// TIA Portal project "ปริญญานิพนธ์" (V17)

(* hardware
DEVICE "S7-1500/ET200MP station_1"  S7-1500 station
   slot 0: "Rail_0"  Rack  6ES7 590-1***0-0AA0
   slot 1: "PLC_1"  CPU 1511-1 PN  6ES7 511-1AK02-0AB0  V2.9
      slot 3: "CPU display_1"  6ES7591-1AA00-0AA0
      slot 32768: "PROFINET interface_1"  X1
         slot 32769: "Port_1"  X1 P1
         slot 32770: "Port_2"  X1 P2
      slot 34817: "Virtual CP interface port_1"  Virtual CP interface port  Virtual CP interface port
DEVICE "HMI_1"  TP900 Comfort
   slot 0: "HMI_1"  TP900 Comfort  6AV2 124-0JC01-0AX0  17.0.0.0
   slot 1: "HMI_RT_1"  TP900 Comfort  6AV2 124-0JC01-0AX0  17.0.0.0
   slot 5: "HMI_1.IE_CP_1"  PROFINET Interface  17.0.0.0
      slot 1: "PROFINET Interface_1"  PROFINET Interface
         slot 1: "Port_1"  Port
         slot 2: "Port_2"  Port
   slot 7: "HMI_1.MPI/DP_CP_1"  MPI/DP Interface  17.0.0.0
*)

// ===== PLC "PLC_1"  CPU 1511-1 PN =====

VAR_GLOBAL   // PLC tag table "Default tag table"
   "ยา 1" AT %MW850 : Word;
   "ยา 2" AT %MW852 : Word;
   "ยา 3" AT %MW854 : Word;
   "ยา 4" AT %MW856 : Word;
   "ยา 5" AT %MW858 : Word;
   "ยา 6" AT %MW860 : Word;
   "ยา 7" AT %MW862 : Word;
   "ยา 8" AT %MW864 : Word;
   "ยา 9" AT %MW866 : Word;
   "ยา 10" AT %MW868 : Word;
   "ยา 11" AT %MW870 : Word;
   "ยา 12" AT %MW872 : Word;
   "ยา 13" AT %MW874 : Word;
   "ยา 14" AT %MW876 : Word;
   "ยา 15" AT %MW878 : Word;
   "ยา 16" AT %MW880 : Word;
   "ยา 17" AT %MW882 : Word;
   "ยา 18" AT %MW884 : Word;
   "ยา 19" AT %MW886 : Word;
   "ยา 20" AT %MW888 : Word;
   "ยา 21" AT %MW890 : Word;
   "ยา 22" AT %MW892 : Word;
   "ยา 23" AT %MW894 : Word;
   "ยา 24" AT %MW896 : Word;
   "ยา 25" AT %MW898 : Word;
   "ยา 26" AT %MW900 : Word;
   "ยา 27" AT %MW902 : Word;
   "ยา 28" AT %MW904 : Word;
   "ยา 29" AT %MW906 : Word;
   "ยา 30" AT %MW908 : Word;
   "ยา 31" AT %MW910 : Word;
   "ยา 32" AT %MW912 : Word;
   "ยา 33" AT %MW914 : Word;
   "ยา 34" AT %MW916 : Word;
   "ยา 35" AT %MW918 : Word;
   "ยา 36" AT %MW920 : Word;
   "ยา 37" AT %MW922 : Word;
   "ยา 38" AT %MW924 : Word;
   "ยา 39" AT %MW926 : Word;
   "ยา 40" AT %MW928 : Word;
   "ยา 41" AT %MW930 : Word;
   "ยา 42" AT %MW932 : Word;
   "ยา 43" AT %MW934 : Word;
   "ยา 44" AT %MW936 : Word;
   "ยา 45" AT %MW938 : Word;
   "ยา 46" AT %MW940 : Word;
   "ยา 47" AT %MW942 : Word;
   "ยา 48" AT %MW944 : Word;
   "ยา 49" AT %MW946 : Word;
   "ยา 50" AT %MW948 : Word;
   "ยา 51" AT %MW950 : Word;
   "ยา 52" AT %MW952 : Word;
   "ยา 53" AT %MW954 : Word;
   "ยา 54" AT %MW956 : Word;
   "ยา 55" AT %MW958 : Word;
   "ยา 56" AT %MW960 : Word;
   "ยา 57" AT %MW962 : Word;
   "ยา 58" AT %MW964 : Word;
   "ยา 59" AT %MW966 : Word;
   "ยา 60" AT %MW968 : Word;
   "ยา 61" AT %MW970 : Word;
   "ยา 62" AT %MW972 : Word;
   "ยา 63" AT %MW974 : Word;
   "ยา 64" AT %MW976 : Word;
   "ยา 65" AT %MW978 : Word;
   "ยา 66" AT %MW980 : Word;
   "ยา 67" AT %MW982 : Word;
   "ยา 68" AT %MW984 : Word;
   "ยา 69" AT %MW986 : Word;
   "ยา 70" AT %MW988 : Word;
   "ยา 71" AT %MW990 : Word;
   "ยา 72" AT %MW992 : Word;
   "ยา 73" AT %MW994 : Word;
   "ยา 74" AT %MW996 : Word;
   "ยา 75" AT %MW998 : Word;
   "ยา 76" AT %MW1000 : Word;
   "ยา 77" AT %MW1002 : Word;
   "ยา 78" AT %MW1004 : Word;
   "ยา 79" AT %MW1006 : Word;
   "ยา 80" AT %MW1008 : Word;
   "ยา 81" AT %MW1010 : Word;
   "ยา 82" AT %MW1012 : Word;
   "ยา 83" AT %MW1014 : Word;
   "ยา 84" AT %MW1016 : Word;
   "ยา 85" AT %MW1018 : Word;
   "ยา 86" AT %MW1020 : Word;
   "ยา 87" AT %MW1022 : Word;
   "ยา 88" AT %MW1024 : Word;
   "ยา 89" AT %MW1026 : Word;
   "ยา 90" AT %MW1028 : Word;
   "ยา 91" AT %MW1030 : Word;
   "ยา 92" AT %MW1032 : Word;
   "ยา 93" AT %MW1034 : Word;
   "ยา 94" AT %MW1036 : Word;
   "ยา 95" AT %MW1038 : Word;
   "ยา 96" AT %MW1040 : Word;
   "ยา 97" AT %MW1042 : Word;
   "ยา 98" AT %MW1044 : Word;
   "ยา 99" AT %MW1046 : Word;
   "ยา 100" AT %MW1048 : Word;
   "ยา 101" AT %MW1050 : Word;
   "ยา 102" AT %MW1052 : Word;
   "ยา 103" AT %MW1054 : Word;
   "ยา 104" AT %MW1056 : Word;
   "ยา 105" AT %MW1058 : Word;
   "ยา 106" AT %MW1060 : Word;
   "ยา 107" AT %MW1062 : Word;
   "ยา 108" AT %MW1064 : Word;
   "ยา 109" AT %MW1066 : Word;
   "ยา 110" AT %MW1068 : Word;
   "ยา 111" AT %MW1070 : Word;
   "ยา 112" AT %MW1072 : Word;
   "ยา 113" AT %MW1074 : Word;
   "ยา 114" AT %MW1076 : Word;
   "ยา 115" AT %MW1078 : Word;
   "ยา 116" AT %MW1080 : Word;
   "ยา 117" AT %MW1082 : Word;
   "ยา 118" AT %MW1084 : Word;
   "ยา 119" AT %MW1086 : Word;
   "ยา 120" AT %MW1088 : Word;
   "ยา 121" AT %MW1090 : Word;
   "ยา 122" AT %MW1092 : Word;
   "ยา 123" AT %MW1094 : Word;
   "ยา 124" AT %MW1096 : Word;
   "ยา 125" AT %MW1098 : Word;
   "ยา 126" AT %MW1100 : Word;
   "ยา 127" AT %MW1102 : Word;
   "ยา 128" AT %MW1104 : Word;
   "ยา 129" AT %MW1106 : Word;
   "ยา 130" AT %MW1108 : Word;
   "ยา 131" AT %MW1110 : Word;
   "ยา 132" AT %MW1112 : Word;
   "ยา 133" AT %MW1114 : Word;
   "ยา 134" AT %MW1116 : Word;
   "ยา 135" AT %MW1118 : Word;
   "ยา 136" AT %MW1120 : Word;
   "ยา 137" AT %MW1122 : Word;
   "ยา 138" AT %MW1124 : Word;
   "ยา 139" AT %MW1126 : Word;
   "ยา 140" AT %MW1128 : Word;
   "ยา 141" AT %MW1130 : Word;
   "ยา 142" AT %MW1132 : Word;
   "ยา 143" AT %MW1134 : Word;
   "ยา 144" AT %MW1136 : Word;
   "ยา 145" AT %MW1138 : Word;
   "ยา 146" AT %MW1140 : Word;
   "ยา 147" AT %MW1142 : Word;
   "ยา 148" AT %MW1144 : Word;
   "ยา 149" AT %MW1146 : Word;
   "ยา 150" AT %MW1148 : Word;
   "ยา 151" AT %MW1150 : Word;
   "ยา 152" AT %MW1152 : Word;
   "ยา 153" AT %MW1154 : Word;
   "ยา 154" AT %MW1156 : Word;
   "ยา 155" AT %MW1158 : Word;
   "ยา 156" AT %MW1160 : Word;
   "ยา 157" AT %MW1162 : Word;
   "ยา 158" AT %MW1164 : Word;
   "ยา 159" AT %MW1166 : Word;
   "ยา 160" AT %MW1168 : Word;
   "ยา 161" AT %MW1170 : Word;
   "ยา 162" AT %MW1172 : Word;
   "ยา 163" AT %MW1174 : Word;
   "\ยา 164" AT %MW1176 : Word;
   "ยา 165" AT %MW1178 : Word;
   "ยา 166" AT %MW1180 : Word;
   "ยา 167" AT %MW1182 : Word;
   "ยา 168" AT %MW1184 : Word;
   "ยา 169" AT %MW1186 : Word;
   "ยา 170" AT %MW1188 : Word;
   "ยา 171" AT %MW1190 : Word;
   "ยา 172" AT %MW1192 : Word;
   "ยา 173" AT %MW1194 : Word;
   "ยา 174" AT %MW1196 : Word;
   "ยา 175" AT %MW1198 : Word;
   "ยา 176" AT %MW1200 : Word;
   "ยา 177" AT %MW1202 : Word;
   "ยา 178" AT %MW1204 : Word;
   "ยา 179" AT %MW1206 : Word;
   "ยา 180" AT %MW1208 : Word;
   "ยา 181" AT %MW1210 : Word;
   "ยา 182" AT %MW1212 : Word;
   "ยา 183" AT %MW1214 : Word;
   "ยา 184" AT %MW1216 : Word;
   "ยา 185" AT %MW1218 : Word;
   "ยา 186" AT %MW1220 : Word;
   "ยา 187" AT %MW1222 : Word;
   "ยา 188" AT %MW1224 : Word;
   "ยา 189" AT %MW1226 : Word;
   "ยา 190" AT %MW1228 : Word;
   "ยา 191" AT %MW1230 : Word;
   "ยา 192" AT %MW1232 : Word;
   "ยา 193" AT %MW1234 : Word;
   "ยา 194" AT %MW1236 : Word;
   "ยา 195" AT %MW1238 : Word;
   "ยา 196" AT %MW1240 : Word;
   "ยา 197" AT %MW1242 : Word;
   "ยา 198" AT %MW1244 : Word;
   "ยา 199" AT %MW1246 : Word;
   "ยา 200" AT %MW1248 : Word;
   "ยา 201" AT %MW1250 : Word;
   "ยา 202" AT %MW1252 : Word;
   "ยา 203" AT %MW1254 : Word;
   "ยา 204" AT %MW1256 : Word;
   "ยา 205" AT %MW1258 : Word;
   "ยา 206" AT %MW1260 : Word;
   "ยา 207" AT %MW1262 : Word;
   "ยา 208" AT %MW1264 : Word;
   "ยา 209" AT %MW1266 : Word;
   "ยา 210" AT %MW1268 : Word;
   "ยา 211" AT %MW1270 : Word;
   "ยา 212" AT %MW1272 : Word;
   "ยา 213" AT %MW1274 : Word;
   "ยา 214" AT %MW1276 : Word;
   "ยา 215" AT %MW1278 : Word;
   "ยา 216" AT %MW1280 : Word;
   "ยา 217" AT %MW1282 : Word;
   "ยา 218" AT %MW1284 : Word;
   "ยา 219" AT %MW1286 : Word;
   "ยา 220" AT %MW1288 : Word;
   "ยา 221" AT %MW1290 : Word;
   "ยา 222" AT %MW1292 : Word;
   "ยา 223" AT %MW1294 : Word;
   "ยา 224" AT %MW1296 : Word;
   "ยา 225" AT %MW1298 : Word;
   "ยา 226" AT %MW1300 : Word;
   "ยา 227" AT %MW1302 : Word;
   "ยา 228" AT %MW1304 : Word;
   "ยา 229" AT %MW1306 : Word;
   "ยา 230" AT %MW1308 : Word;
   "ยา 231" AT %MW1310 : Word;
   "ยา 232" AT %MW1312 : Word;
   "ยา 233" AT %MW1314 : Word;
   "ยา 234" AT %MW1316 : Word;
   "ยา 235" AT %MW1318 : Word;
   "ยา 236" AT %MW1320 : Word;
   "ยา 237" AT %MW1322 : Word;
   "ยา 238" AT %MW1324 : Word;
   "ยา 239" AT %MW1326 : Word;
   "ยา 240" AT %MW1328 : Word;
   "ยา 241" AT %MW1330 : Word;
   "ยา 242" AT %MW1332 : Word;
   "ยา 243" AT %MW1334 : Word;
   "ยา 244" AT %MW1336 : Word;
   "ยา 245" AT %MW1338 : Word;
   "ยา 246" AT %MW1340 : Word;
   "ยา 247" AT %MW1342 : Word;
   "ยา 248" AT %MW1344 : Word;
   "ยา 249" AT %MW1346 : Word;
   "ยา 250" AT %MW1348 : Word;
   "ยา 251" AT %MW1350 : Word;
   "ยา 252" AT %MW1352 : Word;
   "ยา 253" AT %MW1354 : Word;
   "ยา 254" AT %MW1356 : Word;
   "ยา 255" AT %MW1358 : Word;
   "ยา 256" AT %MW1360 : Word;
   "ยา 257" AT %MW1362 : Word;
   "ยา 258" AT %MW1364 : Word;
   "ยา 259" AT %MW1366 : Word;
   "ยา 260" AT %MW1368 : Word;
   "ยา 261" AT %MW1370 : Word;
   "ยา 262" AT %MW1372 : Word;
   "ยา 263" AT %MW1374 : Word;
   "ยา 264" AT %MW1376 : Word;
   "ยา 265" AT %MW1378 : Word;
   "ยา 266" AT %MW1380 : Word;
   "ยา 267" AT %MW1382 : Word;
   "ยา 268" AT %MW1384 : Word;
   "ยา 269" AT %MW1386 : Word;
   "ยา 270" AT %MW1388 : Word;
   "ยา 271" AT %MW1390 : Word;
   "ยา 272" AT %MW1392 : Word;
   "ยา 273" AT %MW1394 : Word;
   "ยา 274" AT %MW1396 : Word;
   "ยา 275" AT %MW1398 : Word;
   "ยา 276" AT %MW1400 : Word;
   "ยา 277" AT %MW1402 : Word;
   "ยา 278" AT %MW1404 : Word;
   "ยา 279" AT %MW1406 : Word;
   "ยา 280" AT %MW1408 : Word;
   "ยา 281" AT %MW1410 : Word;
   "ยา 282" AT %MW1412 : Word;
   "ยา 283" AT %MW1414 : Word;
   "ยา 284" AT %MW1416 : Word;
   "ยา 285" AT %MW1418 : Word;
   "ยา 286" AT %MW1420 : Word;
   "ยา 287" AT %MW1422 : Word;
   "ยา 288" AT %MW1424 : Word;
   "ยา 289" AT %MW1426 : Word;
   "ยา 290" AT %MW1428 : Word;
   "ยา 291" AT %MW1430 : Word;
   "ยา 292" AT %MW1432 : Word;
   "ยา 293" AT %MW1434 : Word;
   "ยา 294" AT %MW1436 : Word;
   "ยา 295" AT %MW1438 : Word;
   "ยา 296" AT %MW1440 : Word;
   "ยา 297" AT %MW1442 : Word;
   "ยา 298" AT %MW1444 : Word;
   "ยา 299" AT %MW1446 : Word;
   "ยา 300" AT %MW1448 : Word;
   "ยา 301" AT %MW1450 : Word;
   "ยา 302" AT %MW1452 : Word;
   "ยา 303" AT %MW1454 : Word;
   "ยา 304" AT %MW1456 : Word;
   "ยา 305" AT %MW1458 : Word;
   "ยา 306" AT %MW1460 : Word;
   "ยา 307" AT %MW1462 : Word;
   "ยา 308" AT %MW1464 : Word;
   "ยา 309" AT %MW1466 : Word;
   "ยา 310" AT %MW1468 : Word;
   "ยา 311" AT %MW1470 : Word;
   "ยา 312" AT %MW1472 : Word;
   "ยา 313" AT %MW1474 : Word;
   "ยา 314" AT %MW1476 : Word;
   "ยา 315" AT %MW1478 : Word;
   "ยา 316" AT %MW1480 : Word;
   "ยา 317" AT %MW1482 : Word;
   "ยา 318" AT %MW1484 : Word;
   "ยา 319" AT %MW1486 : Word;
   "ยา 320" AT %MW1488 : Word;
   "ยา 321" AT %MW1490 : Word;
   "ยา 322" AT %MW1492 : Word;
   "ยา 323" AT %MW1494 : Word;
   "ยา 324" AT %MW1496 : Word;
   "ยา 325" AT %MW1498 : Word;
   "ยา 326" AT %MW1500 : Word;
   "ยา 327" AT %MW1502 : Word;
   "ยา 328" AT %MW1504 : Word;
   "ยา 329" AT %MW1506 : Word;
   "ยา 330" AT %MW1508 : Word;
   "ยา 331" AT %MW1510 : Word;
   "ยา 332" AT %MW1512 : Word;
   "ยา 333" AT %MW1514 : Word;
   "ยา 334" AT %MW1516 : Word;
   "ยา 335" AT %MW1518 : Word;
   "ยา 336" AT %MW1520 : Word;
   "ยา 337" AT %MW1522 : Word;
   "ยา 338" AT %MW1524 : Word;
   "ยา 339" AT %MW1526 : Word;
   "ยา 340" AT %MW1528 : Word;
   "ยา 341" AT %MW1530 : Word;
   "ยา 342" AT %MW1532 : Word;
   "ยา 343" AT %MW1534 : Word;
   "ยา 344" AT %MW1536 : Word;
   "ยา 345" AT %MW1538 : Word;
   "ยา 346" AT %MW1540 : Word;
   "ยา 347" AT %MW1542 : Word;
   "ยา 348" AT %MW1544 : Word;
   "ยา 349" AT %MW1546 : Word;
   "ยา 350" AT %MW1548 : Word;
   "ยา 351" AT %MW1550 : Word;
   "ยา 352" AT %MW1552 : Word;
   "ยา 353" AT %MW1554 : Word;
   "ยา 354" AT %MW1556 : Word;
   "ยา 355" AT %MW1558 : Word;
   "ยา 356" AT %MW1560 : Word;
   "ยา 357" AT %MW1562 : Word;
   "ยา 358" AT %MW1564 : Word;
   "ยา 359" AT %MW1566 : Word;
   "ยา 360" AT %MW1568 : Word;
   "ยา 361" AT %MW1570 : Word;
   "ยา 362" AT %MW1572 : Word;
   "ยา 363" AT %MW1574 : Word;
   "ยา 364" AT %MW1576 : Word;
   "ยา 365" AT %MW1578 : Word;
   "ยา 366" AT %MW1580 : Word;
   "ยา 367" AT %MW1582 : Word;
   "ยา 368" AT %MW1584 : Word;
   "ยา 369" AT %MW1586 : Word;
   "ยา 370" AT %MW1588 : Word;
   "ยา 371" AT %MW1590 : Word;
   "ยา 372" AT %MW1592 : Word;
   "ยา 373" AT %MW1594 : Word;
   "ยา 374" AT %MW1596 : Word;
   "ยา 375" AT %MW1598 : Word;
   "ยา 376" AT %MW1600 : Word;
   "ยา 377" AT %MW1602 : Word;
   "ยา 378" AT %MW1604 : Word;
   "ยา 379" AT %MW1606 : Word;
   "ยา 380" AT %MW1608 : Word;
   "ยา 381" AT %MW1610 : Word;
   "ยา 382" AT %MW1612 : Word;
   "ยา 383" AT %MW1614 : Word;
   "ยา 384" AT %MW1616 : Word;
   "ยา 385" AT %MW1618 : Word;
   "ยา 386" AT %MW1620 : Word;
   "ยา 387" AT %MW1622 : Word;
   "ยา 388" AT %MW1624 : Word;
   "ยา 389" AT %MW1626 : Word;
   "ยา 390" AT %MW1628 : Word;
   "ยา 391" AT %MW1630 : Word;
   "ยา 392" AT %MW1632 : Word;
   "ยา 393" AT %MW1634 : Word;
   "ยา 394" AT %MW1636 : Word;
   "ยา 395" AT %MW1638 : Word;
   "ยา 396" AT %MW1640 : Word;
   "ยา 397" AT %MW1642 : Word;
   "ยา 398" AT %MW1644 : Word;
   "ยา 399" AT %MW1646 : Word;
   "ยา 400" AT %MW1648 : Word;
   "ยา 401" AT %MW1650 : Word;
   "ยา 402" AT %MW1652 : Word;
   "ยา 403" AT %MW1654 : Word;
   "ยา 404" AT %MW1656 : Word;
   "ยา 405" AT %MW1658 : Word;
   "ยา 406" AT %MW1660 : Word;
   "ยา 407" AT %MW1662 : Word;
   "ยา 408" AT %MW1664 : Word;
   "ยา 409" AT %MW1666 : Word;
   "ยา 410" AT %MW1668 : Word;
   "ยา 411" AT %MW1670 : Word;
   "ยา 412" AT %MW1672 : Word;
   "ยา 413" AT %MW1674 : Word;
   "ยา 414" AT %MW1676 : Word;
   "ยา 415" AT %MW1678 : Word;
   "ยา 416" AT %MW1680 : Word;
   "ยา 417" AT %MW1682 : Word;
   "ยา 418" AT %MW1684 : Word;
   "ยา 419" AT %MW1686 : Word;
   "ยา 420" AT %MW1688 : Word;
   "ยา 421" AT %MW1690 : Word;
   "ยา 422" AT %MW1692 : Word;
   "ยา 423" AT %MW1694 : Word;
   "ยา 424" AT %MW1696 : Word;
   "ยา 425" AT %MW1698 : Word;
   "ยา 426" AT %MW1700 : Word;
   "ยา 427" AT %MW1702 : Word;
   "ยา 428" AT %MW1704 : Word;
   "ยา 429" AT %MW1706 : Word;
   "ยา 430" AT %MW1708 : Word;
   "ยา 431" AT %MW1710 : Word;
   "ยา 432" AT %MW1712 : Word;
   "ยา 433" AT %MW1714 : Word;
   "ยา 434" AT %MW1716 : Word;
   "ยา 435" AT %MW1718 : Word;
   "ยา 436" AT %MW1720 : Word;
   "ยา 437" AT %MW1722 : Word;
   "ยา 438" AT %MW1724 : Word;
   "ยา 439" AT %MW1726 : Word;
   "ยา 440" AT %MW1728 : Word;
   "ยา 441" AT %MW1730 : Word;
   "ยา 442" AT %MW1732 : Word;
   "ยา 443" AT %MW1734 : Word;
   "ยา 444" AT %MW1736 : Word;
   "ยา 445" AT %MW1738 : Word;
   "ยา 446" AT %MW1740 : Word;
   "ยา 447" AT %MW1742 : Word;
   "ยา 448" AT %MW1744 : Word;
   "ยา 449" AT %MW1746 : Word;
   "ยา 450" AT %MW1748 : Word;
   "ยา 451" AT %MW1750 : Word;
   "ยา 452" AT %MW1752 : Word;
   "ยา 453" AT %MW1754 : Word;
   "ยา 454" AT %MW1756 : Word;
   "ยา 455" AT %MW1758 : Word;
   "ยา 456" AT %MW1760 : Word;
   "ยา 457" AT %MW1762 : Word;
   "ยา 458" AT %MW1764 : Word;
   "ยา 459" AT %MW1766 : Word;
   "ยา 460" AT %MW1768 : Word;
   "ยา 461" AT %MW1770 : Word;
   "ยา 462" AT %MW1772 : Word;
   "ยา 463" AT %MW1774 : Word;
   "ยา 464" AT %MW1776 : Word;
   "ยา 465" AT %MW1778 : Word;
   "ยา 466" AT %MW1780 : Word;
   "ยา 467" AT %MW1782 : Word;
   "ยา 468" AT %MW1784 : Word;
   "ยา 469" AT %MW1786 : Word;
   "ยา 470" AT %MW1788 : Word;
   "ยา 471" AT %MW1790 : Word;
   "ยา 472" AT %MW1792 : Word;
   "ยา 473" AT %MW1794 : Word;
   "ยา 474" AT %MW1796 : Word;
   "ยา 475" AT %MW1798 : Word;
   "ยา 476" AT %MW1800 : Word;
   "ยา 477" AT %MW1802 : Word;
   "ยา 478" AT %MW1804 : Word;
   "ยา 479" AT %MW1806 : Word;
   "ยา 480" AT %MW1808 : Word;
   "ยา 481" AT %MW1810 : Word;
   "ยา 482" AT %MW1812 : Word;
   "ยา 483" AT %MW1814 : Word;
   "ยา 484" AT %MW1816 : Word;
   "ยา 485" AT %MW1818 : Word;
   "ยา 486" AT %MW1820 : Word;
   "ยา 487" AT %MW1822 : Word;
   "ยา 488" AT %MW1824 : Word;
   "ยา 489" AT %MW1826 : Word;
   "ยา 490" AT %MW1828 : Word;
   "ยา 491" AT %MW1830 : Word;
   "ยา 492" AT %MW1832 : Word;
   "ยา 493" AT %MW1834 : Word;
   "ยา 494" AT %MW1836 : Word;
   "ยา 495" AT %MW1838 : Word;
   "ยา 496" AT %MW1840 : Word;
   "ยา 497" AT %MW1842 : Word;
   "ยา 498" AT %MW1844 : Word;
   "ยา 499" AT %MW1846 : Word;
   "ยา 500" AT %MW1848 : Word;
   "ยา 501" AT %MW1850 : Word;
   "ยา 502" AT %MW1852 : Word;
   "ยา 503" AT %MW1854 : Word;
   "ยา 504" AT %MW1856 : Word;
   "ยา 505" AT %MW1858 : Word;
   "ยา 506" AT %MW1860 : Word;
   "ยา 507" AT %MW1862 : Word;
   "ยา 508" AT %MW1864 : Word;
   "ยา 509" AT %MW1866 : Word;
   "ยา 510" AT %MW1868 : Word;
   "ยา 511" AT %MW1870 : Word;
   "ยา 512" AT %MW1872 : Word;
   "ยา 513" AT %MW1874 : Word;
   "ยา 514" AT %MW1876 : Word;
   "ยา 515" AT %MW1878 : Word;
   "ยา 516" AT %MW1880 : Word;
   "ยา 517" AT %MW1882 : Word;
   "ยา 518" AT %MW1884 : Word;
   "ยา 519" AT %MW1886 : Word;
   "ยา 520" AT %MW1888 : Word;
   "ยา 164" AT %MW1890 : Word;
   "แสดงชื่อยา2" AT %MW3044 : Word;
   "จัดเก็บ Servo DATA 1,2" AT %MW3046 : Word;
   "จัดเก็บ Servo DATA 3" AT %MW3048 : Word;
   "เบิกจ่าย Servo DATA 1,2" AT %MW3050 : Word;
   "เบิกจ่าย Servo DATA 3" AT %MW3052 : Word;
   "Output ปุ่มยืนยันหน้า Screen" AT %M1965.1 : Bool;
   "Output Motor 1,2 fower จัดเก็บ 1" AT %M1892.0 : Bool;
   "Output Motor No3 จัดเก็บ 1" AT %M1892.1 : Bool;
   "หยุดโชว์สถานะมารับยาซ้ำ" AT %M1892.2 : Bool;
   "Output Motor No3 จัดเก็บ 2" AT %M1892.3 : Bool;
   "Output Motor No3จัดเก็บ 3" AT %M1892.4 : Bool;
   "Output Motor No3 จัดเก็บ 4" AT %M1892.5 : Bool;
   "Output Motor No3จัดเก็บ 5" AT %M1892.6 : Bool;
   "Output Motor No3 จัดเก็บ 6" AT %M1892.7 : Bool;
   "Output Motor No3 จัดเก็บ 7" AT %M1893.0 : Bool;
   "Output Motor No3 จัดเก็บ 8" AT %M1893.1 : Bool;
   "Output Motor No3 จัดเก็บ 9" AT %M1893.2 : Bool;
   "Output Motor No3 จัดเก็บ10" AT %M1893.3 : Bool;
   "Output Motor No3จัดเก็บ 11" AT %M1893.4 : Bool;
   "Output Motor No3 จัดเก็บ 12" AT %M1893.5 : Bool;
   "Output Motor No3จัดเก็บ 13" AT %M1893.6 : Bool;
   "Output Motor No3 จัดเก็บ 14" AT %M1893.7 : Bool;
   "Output Motor No3 จัดเก็บ 15" AT %M1894.0 : Bool;
   "Output Motor No3 จัดเก็บ 16" AT %M1894.1 : Bool;
   "Output Motor No3 จัดเก็บ 17" AT %M1894.2 : Bool;
   "Output Motor No3 จัดเก็บ 18" AT %M1894.3 : Bool;
   "Output Motor No3จัดเก็บ 19" AT %M1894.4 : Bool;
   "Output Motor No3 จัดเก็บ 20" AT %M1894.5 : Bool;
   "Output Motor No3จัดเก็บ 21" AT %M1894.6 : Bool;
   "Output Motor No3 จัดเก็บ 22" AT %M1894.7 : Bool;
   "Output Motor No3 จัดเก็บ 23" AT %M1895.0 : Bool;
   "Output Motor No3จัดเก็บ 24" AT %M1895.1 : Bool;
   "Output Motor No3 จัดเก็บ 25" AT %M1895.2 : Bool;
   "Output Motor No3จัดเก็บ 26" AT %M1895.3 : Bool;
   "Oupput Motor 3 จัดเก็บ RESET" AT %M1895.4 : Bool;
   "Output Reset พิเศษ จัดเก็บบ" AT %M1895.5 : Bool;
   "Output Motor 1,2 fower จัดเก็บ 2" AT %M1895.6 : Bool;
   "Output Motor 1,2 fower จัดเก็บ 3" AT %M1895.7 : Bool;
   "Output Motor 1,2 fower จัดเก็บ 4" AT %M1896.0 : Bool;
   "Output Motor 1,2 fower จัดเก็บ 5" AT %M1896.1 : Bool;
   "Output Motor 1,2 fower จัดเก็บ 6" AT %M1896.2 : Bool;
   "Output Motor 1,2 fower จัดเก็บ 7" AT %M1896.3 : Bool;
   "Output Motor 1,2 fower จัดเก็บ 8" AT %M1896.4 : Bool;
   "Output Motor 1,2 fower จัดเก็บ 9" AT %M1896.5 : Bool;
   "Output Motor 1,2 fower จัดเก็บ 10" AT %M1896.6 : Bool;
   "Output Motor 1,2 fower จัดเก็บ 11" AT %M1896.7 : Bool;
   "Output Motor 1,2 fower จัดเก็บ 12" AT %M1897.0 : Bool;
   "Output Motor 1,2 fower จัดเก็บ 13" AT %M1897.1 : Bool;
   "Output Motor 1,2 fower จัดเก็บ 14" AT %M1897.2 : Bool;
   "Output Motor 1,2 fower จัดเก็บ 15" AT %M1897.3 : Bool;
   "Output Motor 1,2 fower จัดเก็บ 16" AT %M1897.4 : Bool;
   "Output Motor 1,2 fower จัดเก็บ 17" AT %M1897.5 : Bool;
   "Output Motor 1,2 fower จัดเก็บ 18" AT %M1897.6 : Bool;
   "Output Motor 1,2 fower จัดเก็บ 19" AT %M1897.7 : Bool;
   "Output Motor 1,2 fower จัดเก็บ 20" AT %M1898.0 : Bool;
   "Output test1" AT %M1898.1 : Bool;
   "Outputtest2" AT %M1898.2 : Bool;
   "Step Motor 3 forword_NOซ้าย-ขวา" AT %M1898.3 : Bool;
   "SR Test" AT %M1898.4 : Bool;
   "Emergency stop" AT %M1898.5 : Bool;
   "Reset-All System" AT %M1898.6 : Bool;
END_VAR

VAR_GLOBAL   // PLC tag table "Tag table_1"
   "SR Conveyor1" AT %M100.0 : Bool;
   "SR Conveyor2" AT %M100.1 : Bool;
   "มีการปุ่มกดยืนยัน" AT %M100.2 : Bool;
   "Brushless Motor Conveyor ทำงาน" AT %M100.3 : Bool;
   "Photoelectic sensor 3 ตรวจเจอวัตถุ" AT %M100.4 : Bool;
   "OutputหลังPhotoelectic sensor 3 ตรวจเจอวัตถุ" AT %M100.5 : Bool;
END_VAR

VAR_GLOBAL   // PLC tag table "Tag table_2"
   "SR_System_In Motor No.1" AT %M200.0 : Bool;
   "SR_System_In Motor No.1(1)" AT %M200.1 : Bool;
   "SR_System_In Motor No.1(2)" AT %M200.2 : Bool;
   "SR_System_In Motor No.1(3)" AT %M200.3 : Bool;
   "SR_System_In Motor No.1(4)" AT %M200.4 : Bool;
   "SR_System_In Motor No.1(5)" AT %M200.5 : Bool;
   "SR_System_In Motor No.1(6)" AT %M200.6 : Bool;
   "SR_System_In Motor No.1(7)" AT %M200.7 : Bool;
   "SR_System_In Motor No.1(8)" AT %M201.0 : Bool;
   "SR_System_In Motor No.1(9)" AT %M201.1 : Bool;
   "SR_System_In Motor No.1(10)" AT %M201.2 : Bool;
   "SR_System_In Motor No.1(11)" AT %M201.3 : Bool;
   "SR_System_In Motor No.1(12)" AT %M201.4 : Bool;
   "SR_System_In Motor No.1(13)" AT %M201.5 : Bool;
   "SR_System_In Motor No.1(14)" AT %M201.6 : Bool;
   "SR_System_In Motor No.1(15)" AT %M201.7 : Bool;
   "SR_System_In Motor No.1(16)" AT %M202.0 : Bool;
   "SR_System_In Motor No.1(17)" AT %M202.1 : Bool;
   "SR_System_In Motor No.1(18)" AT %M202.2 : Bool;
   "SR_System_In Motor No.1(19)" AT %M202.3 : Bool;
   "SR_System_In Motor No.1(20)" AT %M202.4 : Bool;
   "SR_System_In Motor No.1(21)" AT %M202.5 : Bool;
   "SR_System_In Motor No.1(22)" AT %M202.6 : Bool;
   "SR_System_In Motor No.1(23)" AT %M202.7 : Bool;
   "SR_System_In Motor No.1(24)" AT %M203.0 : Bool;
   "SR_System_In Motor No.1(25)" AT %M203.1 : Bool;
   "SR_System_In Motor No.1(26)" AT %M203.2 : Bool;
   "SR_System_In Motor No.1(27)" AT %M203.3 : Bool;
   "SR_System_In Motor No.1(28)" AT %M203.4 : Bool;
   "SR_System_In Motor No.1(29)" AT %M203.5 : Bool;
   "SR_System_In Motor No.1(30)" AT %M203.6 : Bool;
   "SR_System_In Motor No.1(31)" AT %M203.7 : Bool;
   "SR_System_In Motor No.1(32)" AT %M204.0 : Bool;
   "SR_System_In Motor No.1(33)" AT %M204.1 : Bool;
   "SR_System_In Motor No.1(34)" AT %M204.2 : Bool;
   "SR_System_In Motor No.1(35)" AT %M204.3 : Bool;
   "SR_System_In Motor No.1(36)" AT %M204.4 : Bool;
   "SR_System_In Motor No.1(37)" AT %M204.5 : Bool;
   "SR_System_In Motor No.1(38)" AT %M204.6 : Bool;
   "SR_System_In Motor No.1(39)" AT %M204.7 : Bool;
   "Output Step Motor No.1" AT %M205.0 : Bool;
   "Output Step Motor No.2" AT %M205.1 : Bool;
   "Output Step Motor No.3" AT %M205.2 : Bool;
   "Output Step Motor No.4" AT %M205.3 : Bool;
   "Output Step Motor No.5" AT %M205.4 : Bool;
   "Output Step Motor No.6" AT %M205.5 : Bool;
   "Output Step Motor No.7" AT %M205.6 : Bool;
   "Output Step Motor No.8" AT %M205.7 : Bool;
   "Output Step Motor No.9" AT %M206.0 : Bool;
   "Output Step Motor No.10" AT %M206.1 : Bool;
   "Output Step Motor No.11" AT %M206.2 : Bool;
   "Output Step Motor No.12" AT %M206.3 : Bool;
   "Output Step Motor No.13" AT %M206.4 : Bool;
   "Output Step Motor No.14" AT %M206.5 : Bool;
   "Output Step Motor No.15" AT %M206.6 : Bool;
   "Output Step Motor No.16" AT %M206.7 : Bool;
   "Output Step Motor No.17" AT %M207.0 : Bool;
   "Output Step Motor No.18" AT %M207.1 : Bool;
   "Output Step Motor No.19" AT %M207.2 : Bool;
   "Output Step Motor No.20" AT %M207.3 : Bool;
   "Stepper Motor  ทำงาน" AT %M207.4 : Bool;
   "Stepper Motor No.1 ทำงาน" AT %M207.5 : Bool;
   "Stepper Motor No.2 ทำงาน" AT %M207.6 : Bool;
END_VAR

VAR_GLOBAL   // PLC tag table "Tag table_3"
   "Output Step Motor No.31" AT %M300.0 : Bool;
   "SR_System_In Motor No.3.1" AT %M300.1 : Bool;
   "Stepper Motor 3 ทำงาน" AT %M300.2 : Bool;
   "Stepper Motor No.3 ทำงาน" AT %M300.3 : Bool;
   "Outputพิเศษ" AT %M300.4 : Bool;
   "SR สำหรับสั่ง Motor 3 ต่อ1(1)" AT %M300.6 : Bool;
   "SR สำหรับสั่ง Motor 3 ต่อ1(2)" AT %M300.7 : Bool;
   "SR สำหรับสั่ง Motor 3 ต่อ1(3)" AT %M301.0 : Bool;
   "SR สำหรับสั่ง Motor 3 ต่อ1(4)" AT %M301.1 : Bool;
   "SR สำหรับสั่ง Motor 3 ต่อ1(5)" AT %M301.2 : Bool;
   "SR สำหรับสั่ง Motor 3 ต่อ1(6)" AT %M301.3 : Bool;
   "SR สำหรับสั่ง Motor 3 ต่อ1(7)" AT %M301.4 : Bool;
   "SR สำหรับสั่ง Motor 3 ต่อ1(8)" AT %M301.5 : Bool;
   "SR สำหรับสั่ง Motor 3 ต่อ1(9)" AT %M301.6 : Bool;
   "SR สำหรับสั่ง Motor 3 ต่อ1(10)" AT %M301.7 : Bool;
   "SR สำหรับสั่ง Motor 3 ต่อ1(11)" AT %M302.0 : Bool;
   "SR สำหรับสั่ง Motor 3 ต่อ1(12)" AT %M302.1 : Bool;
   "SR สำหรับสั่ง Motor 3 ต่อ1(13)" AT %M302.2 : Bool;
   "SR สำหรับสั่ง Motor 3 ต่อ1(14)" AT %M302.3 : Bool;
   "SR สำหรับสั่ง Motor 3 ต่อ1(15)" AT %M302.4 : Bool;
   "SR สำหรับสั่ง Motor 3 ต่อ1(16)" AT %M302.5 : Bool;
   "SR สำหรับสั่ง Motor 3 ต่อ1(17)" AT %M302.6 : Bool;
   "SR สำหรับสั่ง Motor 3 ต่อ1(18)" AT %M302.7 : Bool;
   "SR สำหรับสั่ง Motor 3 ต่อ1(19)" AT %M303.0 : Bool;
   "SR สำหรับสั่ง Motor 3 ต่อ1(20)" AT %M303.1 : Bool;
   "SR_System_In Motor No.3.2" AT %M300.5 : Bool;
   "SR_System_In Motor No.3.3" AT %M303.2 : Bool;
   "SR_System_In Motor No.3.4" AT %M303.3 : Bool;
   "SR_System_In Motor No.3.5" AT %M303.4 : Bool;
   "SR_System_In Motor No.3.6" AT %M303.5 : Bool;
   "SR_System_In Motor No.3.7" AT %M303.6 : Bool;
   "SR_System_In Motor No.3.8" AT %M303.7 : Bool;
   "SR_System_In Motor No.3.9" AT %M304.0 : Bool;
   "SR_System_In Motor No.3.10" AT %M304.1 : Bool;
   "SR_System_In Motor No.3.11" AT %M304.2 : Bool;
   "SR_System_In Motor No.3.12" AT %M304.3 : Bool;
   "SR_System_In Motor No.3.13" AT %M304.4 : Bool;
   "SR_System_In Motor No.3.14" AT %M304.5 : Bool;
   "SR_System_In Motor No.3.15" AT %M304.6 : Bool;
   "SR_System_In Motor No.3.16" AT %M304.7 : Bool;
   "SR_System_In Motor No.3.17" AT %M305.0 : Bool;
   "SR_System_In Motor No.3.18" AT %M305.1 : Bool;
   "SR_System_In Motor No.3.19" AT %M305.2 : Bool;
   "SR_System_In Motor No.3.20" AT %M305.3 : Bool;
   "SR_System_In Motor No.3.21" AT %M305.4 : Bool;
   "SR_System_In Motor No.3.22" AT %M305.5 : Bool;
   "SR_System_In Motor No.3.23" AT %M305.6 : Bool;
   "SR_System_In Motor No.3.24" AT %M305.7 : Bool;
   "SR_System_In Motor No.3.25" AT %M306.0 : Bool;
   "SR_System_In Motor No.3.26" AT %M306.1 : Bool;
   "Output Step Motor No.32" AT %M306.2 : Bool;
   "Output Step Motor No.33" AT %M306.3 : Bool;
   "Output Step Motor No.34" AT %M306.4 : Bool;
   "Output Step Motor No.35" AT %M306.5 : Bool;
   "Output Step Motor No.36" AT %M306.6 : Bool;
   "Output Step Motor No.37" AT %M306.7 : Bool;
   "Output Step Motor No.38" AT %M307.0 : Bool;
   "Output Step Motor No.39" AT %M307.1 : Bool;
   "Output Step Motor No.40" AT %M307.2 : Bool;
   "Output Step Motor No.41" AT %M307.3 : Bool;
   "Output Step Motor No.42" AT %M307.4 : Bool;
   "Output Step Motor No.43" AT %M307.5 : Bool;
   "Output Step Motor No.44" AT %M307.6 : Bool;
   "Output Step Motor No.45" AT %M307.7 : Bool;
   "Output Step Motor No.46" AT %M308.0 : Bool;
   "Output Step Motor No.47" AT %M308.1 : Bool;
   "Output Step Motor No.48" AT %M308.2 : Bool;
   "Output Step Motor No.49" AT %M308.3 : Bool;
   "Output Step Motor No.50" AT %M308.4 : Bool;
   "Output Step Motor No.51" AT %M308.5 : Bool;
   "Output Step Motor No.52" AT %M308.6 : Bool;
   "Output Step Motor No.53" AT %M308.7 : Bool;
   "Output Step Motor No.54" AT %M309.0 : Bool;
   "Output Step Motor No.55" AT %M309.1 : Bool;
   "Output Step Motor No.56" AT %M309.2 : Bool;
END_VAR

VAR_GLOBAL   // PLC tag table "Tag table_4"
   "Stepper Motor + Gearhead ทำงาน หมุนไปตำแหน่งเริ่มต้น" AT %M400.0 : Bool;
   "Stepper Motor + Gearhead หยุดทำงาน หมุนไปตำแหน่งเริ่มต้น" AT %M400.1 : Bool;
   "Stepper Motor ทำงาน สไลด์ออก" AT %M400.2 : Bool;
   "Stepper Motor หยุดทำงาน สไลด์ออก" AT %M400.3 : Bool;
   "Stepper Motor ทำงาน หนีบกล่องยา" AT %M400.4 : Bool;
   "Stepper Motor หยุดทำงาน หยุดหนหนีบกล่องยา" AT %M400.5 : Bool;
   "Stepper Motor ทำงาน สไลด์เข้า" AT %M400.6 : Bool;
   "Stepper Motor หยุด ทำงานหยุด สไลด์เข้า" AT %M400.7 : Bool;
   "Stepper Motor + Gearhead ทำงาน หมุนไปตำแหน่งทำงานปล่อยกล่องยาลงบนชั้นเก็บกล่องยา" AT %M401.0 : Bool;
   "Stepper Motor + Gearhead หยุดทำงาน หยุดหมุนไปตำแหน่งทำงานปล่อยกล่องยาลงบนชั้นเก็บกล่องยา" AT %M401.1 : Bool;
   "mmตัดการทำงานครบ 1 รอบ" AT %M401.2 : Bool;
   "Stepper Motor ทำงาน ปล่อยกล่องยา" AT %M401.3 : Bool;
   "Stepper Motor หยุด ทำงาน ปล่อยกล่องยา" AT %M401.4 : Bool;
   "SR Gripper No.1" AT %M401.5 : Bool;
   "SR Gripper No.2" AT %M401.6 : Bool;
   "SR Gripper No.3" AT %M401.7 : Bool;
   "SR Gripper No.4" AT %M402.0 : Bool;
   "SR Gripper No.5" AT %M402.1 : Bool;
   "SR Gripper No.6" AT %M402.2 : Bool;
   "SR Gripper No.7" AT %M402.3 : Bool;
   "SR Gripper No.8" AT %M402.4 : Bool;
   "SR Gripper No.9" AT %M402.5 : Bool;
   "Output เมื่อ Motor ถึงตำแหน่งเป้าหมาย" AT %M402.6 : Bool;
   "output Barcoded" AT %M402.7 : Bool;
   "SR Gripper No.10" AT %M403.0 : Bool;
   "หมุนไปตำแหต่งปล่อยกล่องยา" AT %M403.1 : Bool;
END_VAR

VAR_GLOBAL   // PLC tag table "Tag table_5"
   "Blackword SR(1)" AT %M450.0 : Bool;
   "Blackword SR(2)" AT %M450.1 : Bool;
   "Blackword SR(3)" AT %M450.2 : Bool;
   "Blackword SR(4)" AT %M450.3 : Bool;
   "Stepper Motor Blackword  ทำงาน" AT %M450.4 : Bool;
   "Stepper Motor Blackword No.1 ทำงาน" AT %M450.5 : Bool;
   "Stepper Motor Blackword No.2 ทำงาน" AT %M450.6 : Bool;
   "Output Step Motor Blackword  No.1" AT %M450.7 : Bool;
   "Output Step motor  Backword ทำงาน1" AT %M451.0 : Bool;
   "Output Step Motor Blackword  No.2" AT %M451.1 : Bool;
   "Output Step Motor Blackword  No.3" AT %M451.2 : Bool;
   "Output Step Motor Blackword  No.4" AT %M451.3 : Bool;
   "Output Step Motor Blackword  No.5" AT %M451.4 : Bool;
   "Output Step Motor Blackword  No.6" AT %M451.5 : Bool;
   "Output Step Motor Blackword  No.7" AT %M451.6 : Bool;
   "Output Step Motor Blackword  No.8" AT %M451.7 : Bool;
   "Output Step Motor Blackword  No.9" AT %M452.0 : Bool;
   "Output Step Motor Blackword  No.10" AT %M452.1 : Bool;
   "Output Step Motor Blackword  No.11" AT %M452.2 : Bool;
   "Output Step Motor Blackword  No.12" AT %M452.3 : Bool;
   "Output Step Motor Blackword  No.13" AT %M452.4 : Bool;
   "Output Step Motor Blackword  No.14" AT %M452.5 : Bool;
   "Output Step Motor Blackword  No.15" AT %M452.6 : Bool;
   "Output Step Motor Blackword  No.16" AT %M452.7 : Bool;
   "Output Step Motor Blackword  No.17" AT %M453.0 : Bool;
   "Output Step Motor Blackword  No.18" AT %M453.1 : Bool;
   "Output Step Motor Blackword  No.19" AT %M453.2 : Bool;
   "Output Step Motor Blackword  No.20" AT %M453.3 : Bool;
   "Blackword SR(5)" AT %M453.4 : Bool;
   "Blackword SR(6)" AT %M453.5 : Bool;
   "Blackword SR(7)" AT %M453.6 : Bool;
   "Blackword SR(8)" AT %M453.7 : Bool;
   "Blackword SR(9)" AT %M454.0 : Bool;
   "Blackword SR(10)" AT %M454.1 : Bool;
   "Blackword SR(11)" AT %M454.2 : Bool;
   "Blackword SR(12)" AT %M454.3 : Bool;
   "Blackword SR(13)" AT %M454.4 : Bool;
   "Blackword SR(14)" AT %M454.5 : Bool;
   "Blackword SR(15)" AT %M454.6 : Bool;
   "Blackword SR(16)" AT %M454.7 : Bool;
   "Blackword SR(17)" AT %M455.0 : Bool;
   "Blackword SR(18)" AT %M455.1 : Bool;
   "Blackword SR(19)" AT %M455.2 : Bool;
   "Blackword SR(20)" AT %M455.3 : Bool;
   "Blackword SR(21)" AT %M455.4 : Bool;
   "Blackword SR(22)" AT %M455.5 : Bool;
   "Blackword SR(23)" AT %M455.6 : Bool;
   "Blackword SR(24)" AT %M455.7 : Bool;
   "Blackword SR(25)" AT %M456.0 : Bool;
   "Blackword SR(26)" AT %M456.1 : Bool;
   "Blackword SR(27)" AT %M456.2 : Bool;
   "Blackword SR(28)" AT %M456.3 : Bool;
   "Blackword SR(29)" AT %M456.4 : Bool;
   "Blackword SR(30)" AT %M456.5 : Bool;
   "Blackword SR(31)" AT %M456.6 : Bool;
   "Blackword SR(32)" AT %M456.7 : Bool;
   "Blackword SR(33)" AT %M457.0 : Bool;
   "Blackword SR(34)" AT %M457.1 : Bool;
   "Blackword SR(35)" AT %M457.2 : Bool;
   "Blackword SR(36)" AT %M457.3 : Bool;
   "Blackword SR(37)" AT %M457.4 : Bool;
   "Blackword SR(38)" AT %M457.5 : Bool;
   "Blackword SR(39)" AT %M457.6 : Bool;
   "Blackword SR(40)" AT %M457.7 : Bool;
   "Output Step motor  Backword ทำงาน2" AT %M458.0 : Bool;
   "Output Step motor  Backword ทำงาน3" AT %M458.1 : Bool;
   "Output Step motor  Backword ทำงาน4" AT %M458.2 : Bool;
   "Output Step motor  Backword ทำงาน5" AT %M458.3 : Bool;
   "Output Step motor  Backword ทำงาน6" AT %M458.4 : Bool;
   "Output Step motor  Backword ทำงาน7" AT %M458.5 : Bool;
   "Output Step motor  Backword ทำงาน8" AT %M458.6 : Bool;
   "Output Step motor  Backword ทำงาน9" AT %M458.7 : Bool;
   "Output Step motor  Backword ทำงาน10" AT %M459.0 : Bool;
   "Output Step motor  Backword ทำงาน11" AT %M459.1 : Bool;
   "Output Step motor  Backword ทำงาน12" AT %M459.2 : Bool;
   "Output Step motor  Backword ทำงาน13" AT %M459.3 : Bool;
   "Output Step motor  Backword ทำงาน14" AT %M459.4 : Bool;
   "Output Step motor  Backword ทำงาน15" AT %M459.5 : Bool;
   "Output Step motor  Backword ทำงาน16" AT %M459.6 : Bool;
   "Output Step motor  Backword ทำงาน17" AT %M459.7 : Bool;
   "Output Step motor  Backword ทำงาน18" AT %M460.0 : Bool;
   "Output Step motor  Backword ทำงาน19" AT %M460.1 : Bool;
   "Output Step motor  Backword ทำงาน20" AT %M460.2 : Bool;
END_VAR

VAR_GLOBAL   // PLC tag table "Tag table_6"
   "Output Step Motor Blackword  No.1(1)" AT %M550.0 : Bool;
   "SR Step Motor Blackword 1" AT %M550.1 : Bool;
   "SR Step Motor Blackword 2" AT %M550.2 : Bool;
   "Output test1 พิเศษ" AT %M550.7 : Bool;
   "Stepper Motor Blackword3  ทำงาน" AT %M551.0 : Bool;
   "Stepper Motor Blackword No.3 ทำงาน" AT %M551.1 : Bool;
   "output Step motor  Backword ทำงาน No.3(1)" AT %M551.2 : Bool;
   "Output Step Motor Blackword  No.1(2)" AT %M550.3 : Bool;
   "Output Step Motor Blackword  No.1(3)" AT %M550.4 : Bool;
   "Output Step Motor Blackword  No.1(4)" AT %M550.5 : Bool;
   "Output Step Motor Blackword  No.1(5)" AT %M550.6 : Bool;
   "Output Step Motor Blackword  No.1(6)" AT %M551.3 : Bool;
   "Output Step Motor Blackword  No.1(7)" AT %M551.4 : Bool;
   "Output Step Motor Blackword  No.1(8)" AT %M551.5 : Bool;
   "Output Step Motor Blackword  No.1(9)" AT %M551.6 : Bool;
   "Output Step Motor Blackword  No.1(10)" AT %M551.7 : Bool;
   "Output Step Motor Blackword  No.1(11)" AT %M552.0 : Bool;
   "Output Step Motor Blackword  No.1(12)" AT %M552.1 : Bool;
   "Output Step Motor Blackword  No.1(13)" AT %M552.2 : Bool;
   "Output Step Motor Blackword  No.1(14)" AT %M552.3 : Bool;
   "Output Step Motor Blackword  No.1(15)" AT %M552.4 : Bool;
   "Output Step Motor Blackword  No.1(16)" AT %M552.5 : Bool;
   "Output Step Motor Blackword  No.1(17)" AT %M552.6 : Bool;
   "Output Step Motor Blackword  No.1(18)" AT %M552.7 : Bool;
   "Output Step Motor Blackword  No.1(19)" AT %M553.0 : Bool;
   "Output Step Motor Blackword  No.1(20)" AT %M553.1 : Bool;
   "Output Step Motor Blackword  No.1(21)" AT %M553.2 : Bool;
   "Output Step Motor Blackword  No.1(22)" AT %M553.3 : Bool;
   "Output Step Motor Blackword  No.1(23)" AT %M553.4 : Bool;
   "Output Step Motor Blackword  No.1(24)" AT %M553.5 : Bool;
   "Output Step Motor Blackword  No.1(25)" AT %M553.6 : Bool;
   "Output Step Motor Blackword  No.1(26)" AT %M553.7 : Bool;
   "SR Step Motor Blackword 3" AT %M554.0 : Bool;
   "SR Step Motor Blackword 4" AT %M554.1 : Bool;
   "SR Step Motor Blackword 5" AT %M554.2 : Bool;
   "SR Step Motor Blackword 6" AT %M554.3 : Bool;
   "SR Step Motor Blackword 7" AT %M554.4 : Bool;
   "SR Step Motor Blackword 8" AT %M554.5 : Bool;
   "SR Step Motor Blackword 9" AT %M554.6 : Bool;
   "SR Step Motor Blackword 10" AT %M554.7 : Bool;
   "SR Step Motor Blackword 11" AT %M555.0 : Bool;
   "SR Step Motor Blackword 12" AT %M555.1 : Bool;
   "SR Step Motor Blackword 13" AT %M555.2 : Bool;
   "SR Step Motor Blackword 14" AT %M555.3 : Bool;
   "SR Step Motor Blackword 15" AT %M555.4 : Bool;
   "SR Step Motor Blackword 16" AT %M555.5 : Bool;
   "SR Step Motor Blackword 17" AT %M555.6 : Bool;
   "SR Step Motor Blackword 18" AT %M555.7 : Bool;
   "SR Step Motor Blackword 19" AT %M556.0 : Bool;
   "SR Step Motor Blackword 20" AT %M556.1 : Bool;
   "SR Step Motor Blackword 21" AT %M556.2 : Bool;
   "SR Step Motor Blackword 22" AT %M556.3 : Bool;
   "SR Step Motor Blackword 23" AT %M556.4 : Bool;
   "SR Step Motor Blackword 24" AT %M556.5 : Bool;
   "SR Step Motor Blackword 25" AT %M556.6 : Bool;
   "SR Step Motor Blackword 26" AT %M556.7 : Bool;
   "output Step motor  Backword ทำงาน No.3(2)" AT %M557.0 : Bool;
   "output Step motor  Backword ทำงาน No.3(3)" AT %M557.1 : Bool;
   "output Step motor  Backword ทำงาน No.3(4)" AT %M557.2 : Bool;
   "output Step motor  Backword ทำงาน No.3(5)" AT %M557.3 : Bool;
   "output Step motor  Backword ทำงาน No.3(6)" AT %M557.4 : Bool;
   "output Step motor  Backword ทำงาน No.3(7)" AT %M557.5 : Bool;
   "output Step motor  Backword ทำงาน No.3(8)" AT %M557.6 : Bool;
   "output Step motor  Backword ทำงาน No.3(9)" AT %M557.7 : Bool;
   "output Step motor  Backword ทำงาน No.3(10)" AT %M558.0 : Bool;
   "output Step motor  Backword ทำงาน No.3(11)" AT %M558.1 : Bool;
   "output Step motor  Backword ทำงาน No.3(12)" AT %M558.2 : Bool;
   "output Step motor  Backword ทำงาน No.3(13)" AT %M558.3 : Bool;
   "output Step motor  Backword ทำงาน No.3(14)" AT %M558.4 : Bool;
   "output Step motor  Backword ทำงาน No.3(15)" AT %M558.5 : Bool;
   "output Step motor  Backword ทำงาน No.3(16)" AT %M558.6 : Bool;
   "output Step motor  Backword ทำงาน No.3(17)" AT %M558.7 : Bool;
   "output Step motor  Backword ทำงาน No.3(18)" AT %M559.0 : Bool;
   "output Step motor  Backword ทำงาน No.3(19)" AT %M559.1 : Bool;
   "output Step motor  Backword ทำงาน No.3(20)" AT %M559.2 : Bool;
   "output Step motor  Backword ทำงาน No.3(21)" AT %M559.3 : Bool;
   "output Step motor  Backword ทำงาน No.3(22)" AT %M559.4 : Bool;
   "output Step motor  Backword ทำงาน No.3(23)" AT %M559.5 : Bool;
   "output Step motor  Backword ทำงาน No.3(24)" AT %M559.6 : Bool;
   "output Step motor  Backword ทำงาน No.3(25)" AT %M559.7 : Bool;
   "output Step motor  Backword ทำงาน No.3(26)" AT %M560.0 : Bool;
   "SR Step Motor Blackword 27" AT %M560.1 : Bool;
   "SR Step Motor Blackword 28" AT %M560.2 : Bool;
END_VAR

VAR_GLOBAL   // PLC tag table " เบิกจ่าย Forword"
   "SR Step Motro 1,2  เบิกจ่าย 1" AT %M600.0 : Bool;
   "SR Step Motro 1,2  เบิกจ่าย 2" AT %M600.1 : Bool;
   "SR Step Motro 1,2  เบิกจ่าย 3" AT %M600.2 : Bool;
   "SR Step Motro 1,2  เบิกจ่าย 4" AT %M600.3 : Bool;
   "SR Step Motro 1,2  เบิกจ่าย 5" AT %M600.4 : Bool;
   "SR Step Motro 1,2  เบิกจ่าย 6" AT %M600.5 : Bool;
   "SR Step Motro 1,2  เบิกจ่าย 7" AT %M600.6 : Bool;
   "SR Step Motro 1,2  เบิกจ่าย 8" AT %M600.7 : Bool;
   "SR Step Motro 1,2  เบิกจ่าย 9" AT %M601.0 : Bool;
   "SR Step Motro 1,2  เบิกจ่าย 10" AT %M601.1 : Bool;
   "SR Step Motro 1,2  เบิกจ่าย 11" AT %M601.2 : Bool;
   "SR Step Motro 1,2  เบิกจ่าย 12" AT %M601.3 : Bool;
   "SR Step Motro 1,2  เบิกจ่าย 13" AT %M601.4 : Bool;
   "SR Step Motro 1,2  เบิกจ่าย 14" AT %M601.5 : Bool;
   "SR Step Motro 1,2  เบิกจ่าย 15" AT %M601.6 : Bool;
   "SR Step Motro 1,2  เบิกจ่าย 16" AT %M601.7 : Bool;
   "SR Step Motro 1,2  เบิกจ่าย 17" AT %M602.0 : Bool;
   "SR Step Motro 1,2  เบิกจ่าย 18" AT %M602.1 : Bool;
   "SR Step Motro 1,2  เบิกจ่าย 19" AT %M602.2 : Bool;
   "SR Step Motro 1,2  เบิกจ่าย 20" AT %M602.3 : Bool;
   "Outputเมื่อมีการกดปุ่ม 1" AT %M602.4 : Bool;
   "Outputเมื่อมีการกดปุ่ม 2" AT %M602.5 : Bool;
   "Outputเมื่อมีการกดปุ่ม 3" AT %M602.6 : Bool;
   "Outputเมื่อมีการกดปุ่ม 4" AT %M602.7 : Bool;
   "Outputเมื่อมีการกดปุ่ม 5" AT %M603.0 : Bool;
   "Outputเมื่อมีการกดปุ่ม 6" AT %M603.1 : Bool;
   "Outputเมื่อมีการกดปุ่ม 7" AT %M603.2 : Bool;
   "Outputเมื่อมีการกดปุ่ม 8" AT %M603.3 : Bool;
   "Outputเมื่อมีการกดปุ่ม 9" AT %M603.4 : Bool;
   "Outputเมื่อมีการกดปุ่ม 10" AT %M603.5 : Bool;
   "Outputเมื่อมีการกดปุ่ม 11" AT %M603.6 : Bool;
   "Outputเมื่อมีการกดปุ่ม 12" AT %M603.7 : Bool;
   "Outputเมื่อมีการกดปุ่ม 13" AT %M604.0 : Bool;
   "Outputเมื่อมีการกดปุ่ม 14" AT %M604.1 : Bool;
   "Outputเมื่อมีการกดปุ่ม 15" AT %M604.2 : Bool;
   "Outputเมื่อมีการกดปุ่ม 16" AT %M604.3 : Bool;
   "Outputเมื่อมีการกดปุ่ม 17" AT %M604.4 : Bool;
   "Outputเมื่อมีการกดปุ่ม 18" AT %M604.5 : Bool;
   "Outputเมื่อมีการกดปุ่ม 19" AT %M604.6 : Bool;
   "Outputเมื่อมีการกดปุ่ม 20" AT %M604.7 : Bool;
   "Step motor 1,2 NO" AT %M605.0 : Bool;
   "Step motor 1 NO" AT %M605.1 : Bool;
   "Step motor 2 NO" AT %M605.2 : Bool;
   "Output ทำงานเสด M1,2 forword No.1" AT %M605.3 : Bool;
   "Output ทำงานเสด M1,2 forword No.2" AT %M605.4 : Bool;
   "Output ทำงานเสด M1,2 forword No.3" AT %M605.5 : Bool;
   "Output ทำงานเสด M1,2 forword No.4" AT %M605.6 : Bool;
   "Output ทำงานเสด M1,2 forword No.5" AT %M605.7 : Bool;
   "Output ทำงานเสด M1,2 forword No.6" AT %M606.0 : Bool;
   "Output ทำงานเสด M1,2 forword No.7" AT %M606.1 : Bool;
   "Output ทำงานเสด M1,2 forword No.8" AT %M606.2 : Bool;
   "Output ทำงานเสด M1,2 forword No.9" AT %M606.3 : Bool;
   "Output ทำงานเสด M1,2 forword No.10" AT %M606.4 : Bool;
   "Output ทำงานเสด M1,2 forword No.11" AT %M606.5 : Bool;
   "Output ทำงานเสด M1,2 forword No.12" AT %M606.6 : Bool;
   "Output ทำงานเสด M1,2 forword No.13" AT %M606.7 : Bool;
   "Output ทำงานเสด M1,2 forword No.14" AT %M607.0 : Bool;
   "Output ทำงานเสด M1,2 forword No.15" AT %M607.1 : Bool;
   "Output ทำงานเสด M1,2 forword No.16" AT %M607.2 : Bool;
   "Output ทำงานเสด M1,2 forword No.17" AT %M607.3 : Bool;
   "Output ทำงานเสด M1,2 forword No.18" AT %M607.4 : Bool;
   "Output ทำงานเสด M1,2 forword No.19" AT %M607.5 : Bool;
   "Output ทำงานเสด M1,2 forword No.20" AT %M607.6 : Bool;
END_VAR

VAR_GLOBAL   // PLC tag table " เบิกจ่าย Blackword"
   "SR Step Motro 3  เบิกจ่าย 1" AT %M650.0 : Bool;
   "SR Step Motro 3  เบิกจ่าย 2" AT %M650.1 : Bool;
   "SR Step Motro 3  เบิกจ่าย 3" AT %M650.2 : Bool;
   "SR Step Motro 3  เบิกจ่าย 4" AT %M650.3 : Bool;
   "SR Step Motro 3  เบิกจ่าย 5" AT %M650.4 : Bool;
   "SR Step Motro 3  เบิกจ่าย 6" AT %M650.5 : Bool;
   "SR Step Motro 3  เบิกจ่าย 7" AT %M650.6 : Bool;
   "SR Step Motro 3  เบิกจ่าย 8" AT %M650.7 : Bool;
   "SR Step Motro 3  เบิกจ่าย 9" AT %M651.0 : Bool;
   "SR Step Motro 3  เบิกจ่าย 10" AT %M651.1 : Bool;
   "SR Step Motro 3  เบิกจ่าย 11" AT %M651.2 : Bool;
   "SR Step Motro 3  เบิกจ่าย 12" AT %M651.3 : Bool;
   "SR Step Motro 3  เบิกจ่าย 13" AT %M651.4 : Bool;
   "SR Step Motro 3  เบิกจ่าย 14" AT %M651.5 : Bool;
   "SR Step Motro 3  เบิกจ่าย 15" AT %M651.6 : Bool;
   "SR Step Motro 3  เบิกจ่าย 16" AT %M651.7 : Bool;
   "SR Step Motro 3  เบิกจ่าย 17" AT %M652.0 : Bool;
   "SR Step Motro 3  เบิกจ่าย 18" AT %M652.1 : Bool;
   "SR Step Motro 3  เบิกจ่าย 19" AT %M652.2 : Bool;
   "SR Step Motro 3  เบิกจ่าย 20" AT %M652.3 : Bool;
   "output Step motor No.3  1" AT %M652.4 : Bool;
   "output Step motor No.3  2" AT %M652.5 : Bool;
   "output Step motor No.3  3" AT %M652.6 : Bool;
   "output Step motor No.3  4" AT %M652.7 : Bool;
   "output Step motor No.3  5" AT %M653.0 : Bool;
   "output Step motor No.3  6" AT %M653.1 : Bool;
   "output Step motor No.3  7" AT %M653.2 : Bool;
   "output Step motor No.3  8" AT %M653.3 : Bool;
   "output Step motor No.3  9" AT %M653.4 : Bool;
   "output Step motor No.3  10" AT %M653.5 : Bool;
   "output Step motor No.3  11" AT %M653.6 : Bool;
   "output Step motor No.3  12" AT %M653.7 : Bool;
   "output Step motor No.3  13" AT %M654.0 : Bool;
   "output Step motor No.3  14" AT %M654.1 : Bool;
   "output Step motor No.3  15" AT %M654.2 : Bool;
   "output Step motor No.3  16" AT %M654.3 : Bool;
   "output Step motor No.3  17" AT %M654.4 : Bool;
   "output Step motor No.3  18" AT %M654.5 : Bool;
   "output Step motor No.3  19" AT %M654.6 : Bool;
   "output Step motor No.3  20" AT %M654.7 : Bool;
   "Stepper Motor  ทำงาน Blackword_ON" AT %M655.0 : Bool;
   "Step motor 1 Blackword_NO" AT %M655.1 : Bool;
   "Step motor 2 Blackword_NO" AT %M655.2 : Bool;
   "Output No1,2 Blackword 1" AT %M655.3 : Bool;
   "Output No1,2 Blackword 2" AT %M655.4 : Bool;
   "Output No1,2 Blackword 3" AT %M655.5 : Bool;
   "Output No1,2 Blackword 4" AT %M655.6 : Bool;
   "Output No1,2 Blackword 5" AT %M655.7 : Bool;
   "Output No1,2 Blackword 6" AT %M656.0 : Bool;
   "Output No1,2 Blackword 7" AT %M656.1 : Bool;
   "Output No1,2 Blackword 8" AT %M656.2 : Bool;
   "Output No1,2 Blackword 9" AT %M656.3 : Bool;
   "Output No1,2 Blackword 10" AT %M656.4 : Bool;
   "Output No1,2 Blackword 11" AT %M656.5 : Bool;
   "Output No1,2 Blackword 12" AT %M656.6 : Bool;
   "Output No1,2 Blackword 13" AT %M656.7 : Bool;
   "Output No1,2 Blackword 14" AT %M657.0 : Bool;
   "Output No1,2 Blackword 15" AT %M657.1 : Bool;
   "Output No1,2 Blackword 16" AT %M657.2 : Bool;
   "Output No1,2 Blackword 17" AT %M657.3 : Bool;
   "Output No1,2 Blackword 18" AT %M657.4 : Bool;
   "Output No1,2 Blackword 19" AT %M657.5 : Bool;
   "Output No1,2 Blackword 20" AT %M657.6 : Bool;
END_VAR

VAR_GLOBAL   // PLC tag table "Tag table_7"
   "SR  Gripper เบิกจ่าย 1" AT %M700.0 : Bool;
   "SR  Gripper เบิกจ่าย 2" AT %M700.1 : Bool;
   "Output เวลาหลังจากเคลื่ออนที่ไปถึงตำแหน่งเป้าหมาย" AT %M700.2 : Bool;
   "Stepper Motor ทำงาน สไลด์ ตัวงัดกล่องยาออก" AT %M700.3 : Bool;
   "Stepper Motor หยุดทำงาน หยุดสไลด์ ตัวงัดกล่องยาออก" AT %M700.4 : Bool;
   "Stepper Motor ทำงาน สไลด์ ตัวงัดกล่องยาเข้า" AT %M700.5 : Bool;
   "Stepper Motor หยุดทำงาน หยุดสไลด์ ตัวงัดกล่องยาเข้า" AT %M700.6 : Bool;
   "Stepper Motor ทำงาน สั่งconveyor เคลื่อที่ไปข้างหน้า" AT %M700.7 : Bool;
   "Photoelectic Sensor No.1 เบิกจ่าย" AT %M3600.0 : Bool;
   "Photoelectic Sensor No.2 เบิกจ่าย" AT %M3600.1 : Bool;
   "Photoelectic Sensor No.3 เบิกจ่าย" AT %M3600.2 : Bool;
END_VAR

VAR_GLOBAL   // PLC tag table " เบิกจ่าย Blackword 1"
   "SR Blackword Step motor No.3 เบิกจ่าย 1" AT %M800.0 : Bool;
   "SR Blackword Step motor No.3 เบิกจ่าย 2" AT %M800.1 : Bool;
   "SR Blackword Step motor No.3 เบิกจ่าย 3" AT %M800.2 : Bool;
   "SR Blackword Step motor No.3 เบิกจ่าย 4" AT %M800.3 : Bool;
   "SR Blackword Step motor No.3 เบิกจ่าย 5" AT %M800.4 : Bool;
   "SR Blackword Step motor No.3 เบิกจ่าย 6" AT %M800.5 : Bool;
   "SR Blackword Step motor No.3 เบิกจ่าย 7" AT %M800.6 : Bool;
   "SR Blackword Step motor No.3 เบิกจ่าย 8" AT %M800.7 : Bool;
   "SR Blackword Step motor No.3 เบิกจ่าย 9" AT %M801.0 : Bool;
   "SR Blackword Step motor No.3 เบิกจ่าย 10" AT %M801.1 : Bool;
   "SR Blackword Step motor No.3 เบิกจ่าย 11" AT %M801.2 : Bool;
   "SR Blackword Step motor No.3 เบิกจ่าย 12" AT %M801.3 : Bool;
   "SR Blackword Step motor No.3 เบิกจ่าย 13" AT %M801.4 : Bool;
   "SR Blackword Step motor No.3 เบิกจ่าย 14" AT %M801.5 : Bool;
   "SR Blackword Step motor No.3 เบิกจ่าย 15" AT %M801.6 : Bool;
   "SR Blackword Step motor No.3 เบิกจ่าย 16" AT %M801.7 : Bool;
   "SR Blackword Step motor No.3 เบิกจ่าย 17" AT %M802.0 : Bool;
   "SR Blackword Step motor No.3 เบิกจ่าย 18" AT %M802.1 : Bool;
   "SR Blackword Step motor No.3 เบิกจ่าย 19" AT %M802.2 : Bool;
   "SR Blackword Step motor No.3 เบิกจ่าย 20" AT %M802.3 : Bool;
   "SR Blackword Step motor No.3 เบิกจ่าย 21" AT %M802.4 : Bool;
   "SR Blackword Step motor No.3 เบิกจ่าย 22" AT %M802.5 : Bool;
   "SR Blackword Step motor No.3 เบิกจ่าย 23" AT %M802.6 : Bool;
   "SR Blackword Step motor No.3 เบิกจ่าย 24" AT %M802.7 : Bool;
   "SR Blackword Step motor No.3 เบิกจ่าย 25" AT %M803.0 : Bool;
   "SR Blackword Step motor No.3 เบิกจ่าย 26" AT %M803.1 : Bool;
   "Output Blackword Step motor No.3 เบิกจ่าย 1" AT %M803.2 : Bool;
   "Output Blackword Step motor No.3 เบิกจ่าย 2" AT %M803.3 : Bool;
   "Output Blackword Step motor No.3 เบิกจ่าย 3" AT %M803.4 : Bool;
   "Output Blackword Step motor No.3 เบิกจ่าย 4" AT %M803.5 : Bool;
   "Output Blackword Step motor No.3 เบิกจ่าย 5" AT %M803.6 : Bool;
   "Output Blackword Step motor No.3 เบิกจ่าย 6" AT %M803.7 : Bool;
   "Output Blackword Step motor No.3 เบิกจ่าย 7" AT %M804.0 : Bool;
   "Output Blackword Step motor No.3 เบิกจ่าย 8" AT %M804.1 : Bool;
   "Output Blackword Step motor No.3 เบิกจ่าย 9" AT %M804.2 : Bool;
   "Output Blackword Step motor No.3 เบิกจ่าย 10" AT %M804.3 : Bool;
   "Output Blackword Step motor No.3 เบิกจ่าย 11" AT %M804.4 : Bool;
   "Output Blackword Step motor No.3 เบิกจ่าย 12" AT %M804.5 : Bool;
   "Output Blackword Step motor No.3 เบิกจ่าย 13" AT %M804.6 : Bool;
   "Output Blackword Step motor No.3 เบิกจ่าย 14" AT %M804.7 : Bool;
   "Output Blackword Step motor No.3 เบิกจ่าย 15" AT %M805.0 : Bool;
   "Output Blackword Step motor No.3 เบิกจ่าย 16" AT %M805.1 : Bool;
   "Output Blackword Step motor No.3 เบิกจ่าย 17" AT %M805.2 : Bool;
   "Output Blackword Step motor No.3 เบิกจ่าย 18" AT %M805.3 : Bool;
   "Output Blackword Step motor No.3 เบิกจ่าย 19" AT %M805.4 : Bool;
   "Output Blackword Step motor No.3 เบิกจ่าย 20" AT %M805.5 : Bool;
   "Output Blackword Step motor No.3 เบิกจ่าย 21" AT %M805.6 : Bool;
   "Output Blackword Step motor No.3 เบิกจ่าย 22" AT %M805.7 : Bool;
   "Output Blackword Step motor No.3 เบิกจ่าย 23" AT %M806.0 : Bool;
   "Output Blackword Step motor No.3 เบิกจ่าย 24" AT %M806.1 : Bool;
   "Output Blackword Step motor No.3 เบิกจ่าย 25" AT %M806.2 : Bool;
   "Output Blackword Step motor No.3 เบิกจ่าย 26" AT %M806.3 : Bool;
   "เวลาหลังจากเคลื่อนที่ถึงตำแหน่งเป้าหมาย (26) Blackword" AT %M806.4 : Bool;
   "Step Motor 3 Blackword_NO" AT %M806.5 : Bool;
   "Step Motor No.3 Blackword_NO" AT %M806.6 : Bool;
   "Output black No3 1" AT %M806.7 : Bool;
   "Output black No3 2" AT %M807.0 : Bool;
   "Output black No3 3" AT %M807.1 : Bool;
   "Output black No3 4" AT %M807.2 : Bool;
   "Output black No3 5" AT %M807.3 : Bool;
   "Output black No3 6" AT %M807.4 : Bool;
   "Output black No3 7" AT %M807.5 : Bool;
   "Output black No3 8" AT %M807.6 : Bool;
   "Output black No3 9" AT %M807.7 : Bool;
   "Output black No3 10" AT %M808.0 : Bool;
   "Output black No3 11" AT %M808.1 : Bool;
   "Output black No3 12" AT %M808.2 : Bool;
   "Output black No3 13" AT %M808.3 : Bool;
   "Output black No3 14" AT %M808.4 : Bool;
   "Output black No3 15" AT %M808.5 : Bool;
   "Output black No3 16" AT %M808.6 : Bool;
   "Output black No3 17" AT %M808.7 : Bool;
   "Output black No3 18" AT %M809.0 : Bool;
   "Output black No3 19" AT %M809.1 : Bool;
   "Output black No3 20" AT %M809.2 : Bool;
   "Output black No3 21" AT %M809.3 : Bool;
   "Output black No3 22" AT %M809.4 : Bool;
   "Output black No3 23" AT %M809.5 : Bool;
   "Output black No3 24" AT %M809.6 : Bool;
   "Output black No3 25" AT %M809.7 : Bool;
   "Output black No3 26" AT %M810.0 : Bool;
END_VAR

VAR_GLOBAL   // PLC tag table " เบิกจ่าย Forword 1"
   "SR forword Step motor No.3 เบิกจ่าย 1" AT %M750.0 : Bool;
   "SR forword Step motor No.3 เบิกจ่าย 2" AT %M750.1 : Bool;
   "SR forword Step motor No.3 เบิกจ่าย 3" AT %M750.2 : Bool;
   "SR forword Step motor No.3 เบิกจ่าย 4" AT %M750.3 : Bool;
   "SR forword Step motor No.3 เบิกจ่าย 5" AT %M750.4 : Bool;
   "SR forword Step motor No.3 เบิกจ่าย 6" AT %M750.5 : Bool;
   "SR forword Step motor No.3 เบิกจ่าย 7" AT %M750.6 : Bool;
   "SR forword Step motor No.3 เบิกจ่าย 8" AT %M750.7 : Bool;
   "SR forword Step motor No.3 เบิกจ่าย 9" AT %M751.0 : Bool;
   "SR forword Step motor No.3 เบิกจ่าย 10" AT %M751.1 : Bool;
   "SR forword Step motor No.3 เบิกจ่าย 11" AT %M751.2 : Bool;
   "SR forword Step motor No.3 เบิกจ่าย 12" AT %M751.3 : Bool;
   "SR forword Step motor No.3 เบิกจ่าย 13" AT %M751.4 : Bool;
   "SR forword Step motor No.3 เบิกจ่าย 14" AT %M751.5 : Bool;
   "SR forword Step motor No.3 เบิกจ่าย 15" AT %M751.6 : Bool;
   "SR forword Step motor No.3 เบิกจ่าย 16" AT %M751.7 : Bool;
   "SR forword Step motor No.3 เบิกจ่าย 17" AT %M752.0 : Bool;
   "SR forword Step motor No.3 เบิกจ่าย 18" AT %M752.1 : Bool;
   "SR forword Step motor No.3 เบิกจ่าย 19" AT %M752.2 : Bool;
   "SR forword Step motor No.3 เบิกจ่าย 20" AT %M752.3 : Bool;
   "SR forword Step motor No.3 เบิกจ่าย 21" AT %M752.4 : Bool;
   "SR forword Step motor No.3 เบิกจ่าย 22" AT %M752.5 : Bool;
   "SR forword Step motor No.3 เบิกจ่าย 23" AT %M752.6 : Bool;
   "SR forword Step motor No.3 เบิกจ่าย 24" AT %M752.7 : Bool;
   "SR forword Step motor No.3 เบิกจ่าย 25" AT %M753.0 : Bool;
   "SR forword Step motor No.3 เบิกจ่าย 26" AT %M753.1 : Bool;
   "Output forword Step motor No.3 เบิกจ่าย 1" AT %M753.2 : Bool;
   "Output forword Step motor No.3 เบิกจ่าย 2" AT %M753.3 : Bool;
   "Output forword Step motor No.3 เบิกจ่าย 3" AT %M753.4 : Bool;
   "Output forword Step motor No.3 เบิกจ่าย 4" AT %M753.5 : Bool;
   "Output forword Step motor No.3 เบิกจ่าย 5" AT %M753.6 : Bool;
   "Output forword Step motor No.3 เบิกจ่าย 6" AT %M753.7 : Bool;
   "Output forword Step motor No.3 เบิกจ่าย 7" AT %M754.0 : Bool;
   "Output forword Step motor No.3 เบิกจ่าย 8" AT %M754.1 : Bool;
   "Output forword Step motor No.3 เบิกจ่าย 9" AT %M754.2 : Bool;
   "Output forword Step motor No.3 เบิกจ่าย 10" AT %M754.3 : Bool;
   "Output forword Step motor No.3 เบิกจ่าย 11" AT %M754.4 : Bool;
   "Output forword Step motor No.3 เบิกจ่าย 12" AT %M754.5 : Bool;
   "Output forword Step motor No.3 เบิกจ่าย 13" AT %M754.6 : Bool;
   "Output forword Step motor No.3 เบิกจ่าย 14" AT %M754.7 : Bool;
   "Output forword Step motor No.3 เบิกจ่าย 15" AT %M755.0 : Bool;
   "Output forword Step motor No.3 เบิกจ่าย 16" AT %M755.1 : Bool;
   "Output forword Step motor No.3 เบิกจ่าย 17" AT %M755.2 : Bool;
   "Output forword Step motor No.3 เบิกจ่าย 18" AT %M755.3 : Bool;
   "Output forword Step motor No.3 เบิกจ่าย 19" AT %M755.4 : Bool;
   "Output forword Step motor No.3 เบิกจ่าย 20" AT %M755.5 : Bool;
   "Output forword Step motor No.3 เบิกจ่าย 23" AT %M755.6 : Bool;
   "Output forword Step motor No.3 เบิกจ่าย 24" AT %M755.7 : Bool;
   "Output forword Step motor No.3 เบิกจ่าย 25" AT %M756.0 : Bool;
   "Output forword Step motor No.3 เบิกจ่าย 26" AT %M756.1 : Bool;
   "Output forword Step motor No.3 เบิกจ่าย 21" AT %M756.2 : Bool;
   "Output forword Step motor No.3 เบิกจ่าย 22" AT %M756.3 : Bool;
   "เวลาหลังจากเคลื่อนที่ถึงตำแหน่งเป้าหมาย เบิกจ่าย" AT %M756.4 : Bool;
   "Step Motor 3 forword_NO" AT %M756.5 : Bool;
   "Step Motor No.3 forword_NO" AT %M756.6 : Bool;
   "SR หลังจาก Motor 1,2 ทำงานเสด" AT %M756.7 : Bool;
   "Output ทำงานเสด M 3 forword No.1" AT %M757.0 : Bool;
   "Output ทำงานเสด M 3 forword No.2" AT %M757.1 : Bool;
   "Output ทำงานเสด M 3 forword No.3" AT %M757.2 : Bool;
   "Output ทำงานเสด M 3 forword No.4" AT %M757.3 : Bool;
   "Output ทำงานเสด M 3 forword No.5" AT %M757.4 : Bool;
   "Output ทำงานเสด M 3 forword No.6" AT %M757.5 : Bool;
   "Output ทำงานเสด M 3 forword No.7" AT %M757.6 : Bool;
   "Output ทำงานเสด M 3 forword No.8" AT %M757.7 : Bool;
   "Output ทำงานเสด M 3 forword No.9" AT %M758.0 : Bool;
   "Output ทำงานเสด M 3 forword No.10" AT %M758.1 : Bool;
   "Output ทำงานเสด M 3 forword No.11" AT %M758.2 : Bool;
   "Output ทำงานเสด M 3 forword No.12" AT %M758.3 : Bool;
   "Output ทำงานเสด M 3 forword No.13" AT %M758.4 : Bool;
   "Output ทำงานเสด M 3 forword No.14" AT %M758.5 : Bool;
   "Output ทำงานเสด M 3 forword No.15" AT %M758.6 : Bool;
   "Output ทำงานเสด M 3 forword No.16" AT %M758.7 : Bool;
   "Output ทำงานเสด M 3 forword No.17" AT %M759.0 : Bool;
   "Output ทำงานเสด M 3 forword No.18" AT %M759.1 : Bool;
   "Output ทำงานเสด M 3 forword No.19" AT %M759.2 : Bool;
   "Output ทำงานเสด M 3 forword No.20" AT %M759.3 : Bool;
   "Output ทำงานเสด M 3 forword No.21" AT %M759.4 : Bool;
   "Output ทำงานเสด M 3 forword No.22" AT %M759.5 : Bool;
   "Output ทำงานเสด M 3 forword No.23" AT %M759.6 : Bool;
   "Output ทำงานเสด M 3 forword No.24" AT %M759.7 : Bool;
   "Output ทำงานเสด M 3 forword No.25" AT %M760.0 : Bool;
   "Output ทำงานเสด M 3 forword No.26" AT %M760.1 : Bool;
END_VAR

VAR_GLOBAL   // PLC tag table "Tag table_8"
   "M1" AT %M1900.0 : Bool;
   "M2" AT %M1900.1 : Bool;
   "M3" AT %M1900.2 : Bool;
   "M4" AT %M1900.3 : Bool;
   "M5" AT %M1900.4 : Bool;
   "M6" AT %M1900.5 : Bool;
   "M7" AT %M1900.6 : Bool;
   "M8" AT %M1900.7 : Bool;
   "M9" AT %M1901.0 : Bool;
   "M10" AT %M1901.1 : Bool;
   "M11" AT %M1901.2 : Bool;
   "M12" AT %M1901.3 : Bool;
   "M13" AT %M1901.4 : Bool;
   "M14" AT %M1901.5 : Bool;
   "M15" AT %M1901.6 : Bool;
   "M16" AT %M1901.7 : Bool;
   "M17" AT %M1902.0 : Bool;
   "M18" AT %M1902.1 : Bool;
   "M19" AT %M1902.2 : Bool;
   "M20" AT %M1902.3 : Bool;
   "M21" AT %M1902.4 : Bool;
   "M22" AT %M1902.5 : Bool;
   "M23" AT %M1902.6 : Bool;
   "M24" AT %M1902.7 : Bool;
   "M25" AT %M1903.0 : Bool;
   "M26" AT %M1903.1 : Bool;
   "M27" AT %M1903.2 : Bool;
   "M28" AT %M1903.3 : Bool;
   "M29" AT %M1903.4 : Bool;
   "M30" AT %M1903.5 : Bool;
   "M31" AT %M1903.6 : Bool;
   "M32" AT %M1903.7 : Bool;
   "M33" AT %M1904.0 : Bool;
   "M34" AT %M1904.1 : Bool;
   "M35" AT %M1904.2 : Bool;
   "M36" AT %M1904.3 : Bool;
   "M37" AT %M1904.4 : Bool;
   "M38" AT %M1904.5 : Bool;
   "M39" AT %M1904.6 : Bool;
   "M40" AT %M1904.7 : Bool;
   "M41" AT %M1905.0 : Bool;
   "M42" AT %M1905.1 : Bool;
   "M43" AT %M1905.2 : Bool;
   "M44" AT %M1905.3 : Bool;
   "M45" AT %M1905.4 : Bool;
   "M46" AT %M1905.5 : Bool;
   "M47" AT %M1905.6 : Bool;
   "M48" AT %M1905.7 : Bool;
   "M49" AT %M1906.0 : Bool;
   "M50" AT %M1906.1 : Bool;
   "M51" AT %M1906.2 : Bool;
   "M52" AT %M1906.3 : Bool;
   "M53" AT %M1906.4 : Bool;
   "M54" AT %M1906.5 : Bool;
   "M55" AT %M1906.6 : Bool;
   "M56" AT %M1906.7 : Bool;
   "M57" AT %M1907.0 : Bool;
   "M58" AT %M1907.1 : Bool;
   "M59" AT %M1907.2 : Bool;
   "M60" AT %M1907.3 : Bool;
   "M61" AT %M1907.4 : Bool;
   "M62" AT %M1907.5 : Bool;
   "M63" AT %M1907.6 : Bool;
   "M64" AT %M1907.7 : Bool;
   "M65" AT %M1908.0 : Bool;
   "M66" AT %M1908.1 : Bool;
   "M67" AT %M1908.2 : Bool;
   "M68" AT %M1908.3 : Bool;
   "M69" AT %M1908.4 : Bool;
   "M70" AT %M1908.5 : Bool;
   "M71" AT %M1908.6 : Bool;
   "M72" AT %M1908.7 : Bool;
   "M73" AT %M1909.0 : Bool;
   "M74" AT %M1909.1 : Bool;
   "M75" AT %M1909.2 : Bool;
   "M76" AT %M1909.3 : Bool;
   "M77" AT %M1909.4 : Bool;
   "M78" AT %M1909.5 : Bool;
   "M79" AT %M1909.6 : Bool;
   "M80" AT %M1909.7 : Bool;
   "M81" AT %M1910.0 : Bool;
   "M82" AT %M1910.1 : Bool;
   "M83" AT %M1910.2 : Bool;
   "M84" AT %M1910.3 : Bool;
   "M85" AT %M1910.4 : Bool;
   "M86" AT %M1910.5 : Bool;
   "M87" AT %M1910.6 : Bool;
   "M88" AT %M1910.7 : Bool;
   "M89" AT %M1911.0 : Bool;
   "M90" AT %M1911.1 : Bool;
   "M91" AT %M1911.2 : Bool;
   "M92" AT %M1911.3 : Bool;
   "M93" AT %M1911.4 : Bool;
   "M94" AT %M1911.5 : Bool;
   "M95" AT %M1911.6 : Bool;
   "M96" AT %M1911.7 : Bool;
   "M97" AT %M1912.0 : Bool;
   "M98" AT %M1912.1 : Bool;
   "M99" AT %M1912.2 : Bool;
   "M100" AT %M1912.3 : Bool;
   "M101" AT %M1912.4 : Bool;
   "M102" AT %M1912.5 : Bool;
   "M103" AT %M1912.6 : Bool;
   "M104" AT %M1912.7 : Bool;
   "M105" AT %M1913.0 : Bool;
   "M106" AT %M1913.1 : Bool;
   "M107" AT %M1913.2 : Bool;
   "M108" AT %M1913.3 : Bool;
   "M109" AT %M1913.4 : Bool;
   "M110" AT %M1913.5 : Bool;
   "M111" AT %M1913.6 : Bool;
   "M112" AT %M1913.7 : Bool;
   "M113" AT %M1914.0 : Bool;
   "M114" AT %M1914.1 : Bool;
   "M115" AT %M1914.2 : Bool;
   "M116" AT %M1914.3 : Bool;
   "M117" AT %M1914.4 : Bool;
   "M118" AT %M1914.5 : Bool;
   "M119" AT %M1914.6 : Bool;
   "M120" AT %M1914.7 : Bool;
   "M121" AT %M1915.0 : Bool;
   "M122" AT %M1915.1 : Bool;
   "M123" AT %M1915.2 : Bool;
   "M124" AT %M1915.3 : Bool;
   "M125" AT %M1915.4 : Bool;
   "M126" AT %M1915.5 : Bool;
   "M127" AT %M1915.6 : Bool;
   "M128" AT %M1915.7 : Bool;
   "M129" AT %M1916.0 : Bool;
   "M130" AT %M1916.1 : Bool;
   "M131" AT %M1916.2 : Bool;
   "M132" AT %M1916.3 : Bool;
   "M133" AT %M1916.4 : Bool;
   "M134" AT %M1916.5 : Bool;
   "M135" AT %M1916.6 : Bool;
   "M136" AT %M1916.7 : Bool;
   "M137" AT %M1917.0 : Bool;
   "M138" AT %M1917.1 : Bool;
   "M139" AT %M1917.2 : Bool;
   "M140" AT %M1917.3 : Bool;
   "M141" AT %M1917.4 : Bool;
   "M142" AT %M1917.5 : Bool;
   "M143" AT %M1917.6 : Bool;
   "M144" AT %M1917.7 : Bool;
   "M145" AT %M1918.0 : Bool;
   "M146" AT %M1918.1 : Bool;
   "M147" AT %M1918.2 : Bool;
   "M148" AT %M1918.3 : Bool;
   "M149" AT %M1918.4 : Bool;
   "M150" AT %M1918.5 : Bool;
   "M151" AT %M1918.6 : Bool;
   "M152" AT %M1918.7 : Bool;
   "M153" AT %M1919.0 : Bool;
   "M154" AT %M1919.1 : Bool;
   "M155" AT %M1919.2 : Bool;
   "M156" AT %M1919.3 : Bool;
   "M157" AT %M1919.4 : Bool;
   "M158" AT %M1919.5 : Bool;
   "M159" AT %M1919.6 : Bool;
   "M160" AT %M1919.7 : Bool;
   "M161" AT %M1920.0 : Bool;
   "M162" AT %M1920.1 : Bool;
   "M163" AT %M1920.2 : Bool;
   "M164" AT %M1920.3 : Bool;
   "M165" AT %M1920.4 : Bool;
   "M166" AT %M1920.5 : Bool;
   "M167" AT %M1920.6 : Bool;
   "M168" AT %M1920.7 : Bool;
   "M169" AT %M1921.0 : Bool;
   "M170" AT %M1921.1 : Bool;
   "M171" AT %M1921.2 : Bool;
   "M172" AT %M1921.3 : Bool;
   "M173" AT %M1921.4 : Bool;
   "M174" AT %M1921.5 : Bool;
   "M175" AT %M1921.6 : Bool;
   "M176" AT %M1921.7 : Bool;
   "M177" AT %M1922.0 : Bool;
   "M178" AT %M1922.1 : Bool;
   "M179" AT %M1922.2 : Bool;
   "M180" AT %M1922.3 : Bool;
   "M181" AT %M1922.4 : Bool;
   "M182" AT %M1922.5 : Bool;
   "M183" AT %M1922.6 : Bool;
   "M184" AT %M1922.7 : Bool;
   "M185" AT %M1923.0 : Bool;
   "M186" AT %M1923.1 : Bool;
   "M187" AT %M1923.2 : Bool;
   "M188" AT %M1923.3 : Bool;
   "M189" AT %M1923.4 : Bool;
   "M190" AT %M1923.5 : Bool;
   "M191" AT %M1923.6 : Bool;
   "M192" AT %M1923.7 : Bool;
   "M193" AT %M1924.0 : Bool;
   "M194" AT %M1924.1 : Bool;
   "M195" AT %M1924.2 : Bool;
   "M196" AT %M1924.3 : Bool;
   "M197" AT %M1924.4 : Bool;
   "M198" AT %M1924.5 : Bool;
   "M199" AT %M1924.6 : Bool;
   "M200" AT %M1924.7 : Bool;
   "M201" AT %M1925.0 : Bool;
   "M202" AT %M1925.1 : Bool;
   "M203" AT %M1925.2 : Bool;
   "M204" AT %M1925.3 : Bool;
   "M205" AT %M1925.4 : Bool;
   "M206" AT %M1925.5 : Bool;
   "M207" AT %M1925.6 : Bool;
   "M208" AT %M1925.7 : Bool;
   "M209" AT %M1926.0 : Bool;
   "M210" AT %M1926.1 : Bool;
   "M211" AT %M1926.2 : Bool;
   "M212" AT %M1926.3 : Bool;
   "M213" AT %M1926.4 : Bool;
   "M214" AT %M1926.5 : Bool;
   "M215" AT %M1926.6 : Bool;
   "M216" AT %M1926.7 : Bool;
   "M217" AT %M1927.0 : Bool;
   "M218" AT %M1927.1 : Bool;
   "M219" AT %M1927.2 : Bool;
   "M220" AT %M1927.3 : Bool;
   "M221" AT %M1927.4 : Bool;
   "M222" AT %M1927.5 : Bool;
   "M223" AT %M1927.6 : Bool;
   "M224" AT %M1927.7 : Bool;
   "M225" AT %M1928.0 : Bool;
   "M226" AT %M1928.1 : Bool;
   "M227" AT %M1928.2 : Bool;
   "M228" AT %M1928.3 : Bool;
   "M229" AT %M1928.4 : Bool;
   "M230" AT %M1928.5 : Bool;
   "M231" AT %M1928.6 : Bool;
   "M232" AT %M1928.7 : Bool;
   "M233" AT %M1929.0 : Bool;
   "M234" AT %M1929.1 : Bool;
   "M235" AT %M1929.2 : Bool;
   "M236" AT %M1929.3 : Bool;
   "M237" AT %M1929.4 : Bool;
   "M238" AT %M1929.5 : Bool;
   "M239" AT %M1929.6 : Bool;
   "M240" AT %M1929.7 : Bool;
   "M241" AT %M1930.0 : Bool;
   "M242" AT %M1930.1 : Bool;
   "M243" AT %M1930.2 : Bool;
   "M244" AT %M1930.3 : Bool;
   "M245" AT %M1930.4 : Bool;
   "M246" AT %M1930.5 : Bool;
   "M247" AT %M1930.6 : Bool;
   "M248" AT %M1930.7 : Bool;
   "M249" AT %M1931.0 : Bool;
   "M250" AT %M1931.1 : Bool;
   "M251" AT %M1931.2 : Bool;
   "M252" AT %M1931.3 : Bool;
   "M253" AT %M1931.4 : Bool;
   "M254" AT %M1931.5 : Bool;
   "M255" AT %M1931.6 : Bool;
   "M256" AT %M1931.7 : Bool;
   "M257" AT %M1932.0 : Bool;
   "M258" AT %M1932.1 : Bool;
   "M259" AT %M1932.2 : Bool;
   "M260" AT %M1932.3 : Bool;
   "M261" AT %M1932.4 : Bool;
   "M262" AT %M1932.5 : Bool;
   "M263" AT %M1932.6 : Bool;
   "M264" AT %M1932.7 : Bool;
   "M265" AT %M1933.0 : Bool;
   "M266" AT %M1933.1 : Bool;
   "M267" AT %M1933.2 : Bool;
   "M268" AT %M1933.3 : Bool;
   "M269" AT %M1933.4 : Bool;
   "M270" AT %M1933.5 : Bool;
   "M271" AT %M1933.6 : Bool;
   "M272" AT %M1933.7 : Bool;
   "M273" AT %M1934.0 : Bool;
   "M274" AT %M1934.1 : Bool;
   "M275" AT %M1934.2 : Bool;
   "M276" AT %M1934.3 : Bool;
   "M277" AT %M1934.4 : Bool;
   "M278" AT %M1934.5 : Bool;
   "M279" AT %M1934.6 : Bool;
   "M280" AT %M1934.7 : Bool;
   "M281" AT %M1935.0 : Bool;
   "M282" AT %M1935.1 : Bool;
   "M283" AT %M1935.2 : Bool;
   "M284" AT %M1935.3 : Bool;
   "M285" AT %M1935.4 : Bool;
   "M286" AT %M1935.5 : Bool;
   "M287" AT %M1935.6 : Bool;
   "M288" AT %M1935.7 : Bool;
   "M289" AT %M1936.0 : Bool;
   "M290" AT %M1936.1 : Bool;
   "M291" AT %M1936.2 : Bool;
   "M292" AT %M1936.3 : Bool;
   "M294" AT %M1936.4 : Bool;
   "M293" AT %M1936.5 : Bool;
   "M295" AT %M1936.6 : Bool;
   "M296" AT %M1936.7 : Bool;
   "M297" AT %M1937.0 : Bool;
   "M298" AT %M1937.1 : Bool;
   "M299" AT %M1937.2 : Bool;
   "M300" AT %M1937.3 : Bool;
   "M301" AT %M1937.4 : Bool;
   "M302" AT %M1937.5 : Bool;
   "M303" AT %M1937.6 : Bool;
   "M304" AT %M1937.7 : Bool;
   "M305" AT %M1938.0 : Bool;
   "M306" AT %M1938.1 : Bool;
   "M307" AT %M1938.2 : Bool;
   "M308" AT %M1938.3 : Bool;
   "M309" AT %M1938.4 : Bool;
   "M310" AT %M1938.5 : Bool;
   "M311" AT %M1938.6 : Bool;
   "M312" AT %M1938.7 : Bool;
   "M313" AT %M1939.0 : Bool;
   "M314" AT %M1939.1 : Bool;
   "M315" AT %M1939.2 : Bool;
   "M316" AT %M1939.3 : Bool;
   "M317" AT %M1939.4 : Bool;
   "M318" AT %M1939.5 : Bool;
   "M319" AT %M1939.6 : Bool;
   "M320" AT %M1939.7 : Bool;
   "M321" AT %M1940.0 : Bool;
   "M322" AT %M1940.1 : Bool;
   "M323" AT %M1940.2 : Bool;
   "M324" AT %M1940.3 : Bool;
   "M325" AT %M1940.4 : Bool;
   "M326" AT %M1940.5 : Bool;
   "M327" AT %M1940.6 : Bool;
   "M328" AT %M1940.7 : Bool;
   "M329" AT %M1941.0 : Bool;
   "M330" AT %M1941.1 : Bool;
   "M331" AT %M1941.2 : Bool;
   "M332" AT %M1941.3 : Bool;
   "M333" AT %M1941.4 : Bool;
   "M334" AT %M1941.5 : Bool;
   "M335" AT %M1941.6 : Bool;
   "M336" AT %M1941.7 : Bool;
   "M337" AT %M1942.0 : Bool;
   "M338" AT %M1942.1 : Bool;
   "M339" AT %M1942.2 : Bool;
   "M340" AT %M1942.3 : Bool;
   "M341" AT %M1942.4 : Bool;
   "M342" AT %M1942.5 : Bool;
   "M343" AT %M1942.6 : Bool;
   "M344" AT %M1942.7 : Bool;
   "M345" AT %M1943.0 : Bool;
   "M346" AT %M1943.1 : Bool;
   "M347" AT %M1943.2 : Bool;
   "M348" AT %M1943.3 : Bool;
   "M349" AT %M1943.4 : Bool;
   "M350" AT %M1943.5 : Bool;
   "M351" AT %M1943.6 : Bool;
   "M352" AT %M1943.7 : Bool;
   "M353" AT %M1944.0 : Bool;
   "M354" AT %M1944.1 : Bool;
   "M355" AT %M1944.2 : Bool;
   "M356" AT %M1944.3 : Bool;
   "M357" AT %M1944.4 : Bool;
   "M358" AT %M1944.5 : Bool;
   "M359" AT %M1944.6 : Bool;
   "M360" AT %M1944.7 : Bool;
   "M361" AT %M1945.0 : Bool;
   "M362" AT %M1945.1 : Bool;
   "M363" AT %M1945.2 : Bool;
   "M364" AT %M1945.3 : Bool;
   "M365" AT %M1945.4 : Bool;
   "M366" AT %M1945.5 : Bool;
   "M367" AT %M1945.6 : Bool;
   "M368" AT %M1945.7 : Bool;
   "M369" AT %M1946.0 : Bool;
   "M370" AT %M1946.1 : Bool;
   "M371" AT %M1946.2 : Bool;
   "M372" AT %M1946.3 : Bool;
   "M373" AT %M1946.4 : Bool;
   "M374" AT %M1946.5 : Bool;
   "M375" AT %M1946.6 : Bool;
   "M376" AT %M1946.7 : Bool;
   "M377" AT %M1947.0 : Bool;
   "M378" AT %M1947.1 : Bool;
   "M379" AT %M1947.2 : Bool;
   "M380" AT %M1947.3 : Bool;
   "M381" AT %M1947.4 : Bool;
   "M382" AT %M1947.5 : Bool;
   "M383" AT %M1947.6 : Bool;
   "M384" AT %M1947.7 : Bool;
   "M385" AT %M1948.0 : Bool;
   "M386" AT %M1948.1 : Bool;
   "M387" AT %M1948.2 : Bool;
   "M388" AT %M1948.3 : Bool;
   "M389" AT %M1948.4 : Bool;
   "M390" AT %M1948.5 : Bool;
   "M391" AT %M1948.6 : Bool;
   "M392" AT %M1948.7 : Bool;
   "M393" AT %M1949.0 : Bool;
   "M394" AT %M1949.1 : Bool;
   "M395" AT %M1949.2 : Bool;
   "M396" AT %M1949.3 : Bool;
   "M397" AT %M1949.4 : Bool;
   "M398" AT %M1949.5 : Bool;
   "M399" AT %M1949.6 : Bool;
   "M400" AT %M1949.7 : Bool;
   "M401" AT %M1950.0 : Bool;
   "M402" AT %M1950.1 : Bool;
   "M403" AT %M1950.2 : Bool;
   "M404" AT %M1950.3 : Bool;
   "M405" AT %M1950.4 : Bool;
   "M406" AT %M1950.5 : Bool;
   "M407" AT %M1950.6 : Bool;
   "M408" AT %M1950.7 : Bool;
   "M409" AT %M1951.0 : Bool;
   "M410" AT %M1951.1 : Bool;
   "M411" AT %M1951.2 : Bool;
   "M412" AT %M1951.3 : Bool;
   "M413" AT %M1951.4 : Bool;
   "M414" AT %M1951.5 : Bool;
   "M415" AT %M1951.6 : Bool;
   "M416" AT %M1951.7 : Bool;
   "M417" AT %M1952.0 : Bool;
   "M418" AT %M1952.1 : Bool;
   "M419" AT %M1952.2 : Bool;
   "M420" AT %M1952.3 : Bool;
   "M421" AT %M1952.4 : Bool;
   "M422" AT %M1952.5 : Bool;
   "M423" AT %M1952.6 : Bool;
   "M424" AT %M1952.7 : Bool;
   "M425" AT %M1953.0 : Bool;
   "M426" AT %M1953.1 : Bool;
   "M427" AT %M1953.2 : Bool;
   "M428" AT %M1953.3 : Bool;
   "M429" AT %M1953.4 : Bool;
   "M430" AT %M1953.5 : Bool;
   "M431" AT %M1953.6 : Bool;
   "M432" AT %M1953.7 : Bool;
   "M433" AT %M1954.0 : Bool;
   "M434" AT %M1954.1 : Bool;
   "M435" AT %M1954.2 : Bool;
   "M436" AT %M1954.3 : Bool;
   "M437" AT %M1954.4 : Bool;
   "M438" AT %M1954.5 : Bool;
   "M439" AT %M1954.6 : Bool;
   "M440" AT %M1954.7 : Bool;
   "M441" AT %M1955.0 : Bool;
   "M442" AT %M1955.1 : Bool;
   "M443" AT %M1955.2 : Bool;
   "M444" AT %M1955.3 : Bool;
   "M445" AT %M1955.4 : Bool;
   "M446" AT %M1955.5 : Bool;
   "M447" AT %M1955.6 : Bool;
   "M448" AT %M1955.7 : Bool;
   "M449" AT %M1956.0 : Bool;
   "M450" AT %M1956.1 : Bool;
   "M451" AT %M1956.2 : Bool;
   "M452" AT %M1956.3 : Bool;
   "M453" AT %M1956.4 : Bool;
   "M454" AT %M1956.5 : Bool;
   "M455" AT %M1956.6 : Bool;
   "M456" AT %M1956.7 : Bool;
   "M457" AT %M1957.0 : Bool;
   "M458" AT %M1957.1 : Bool;
   "M459" AT %M1957.2 : Bool;
   "M460" AT %M1957.3 : Bool;
   "M461" AT %M1957.4 : Bool;
   "M462" AT %M1957.5 : Bool;
   "M463" AT %M1957.6 : Bool;
   "M464" AT %M1957.7 : Bool;
   "M465" AT %M1958.0 : Bool;
   "M466" AT %M1958.1 : Bool;
   "M467" AT %M1958.2 : Bool;
   "M468" AT %M1958.3 : Bool;
   "M469" AT %M1958.4 : Bool;
   "M470" AT %M1958.5 : Bool;
   "M471" AT %M1958.6 : Bool;
   "M472" AT %M1958.7 : Bool;
   "M473" AT %M1959.0 : Bool;
   "M474" AT %M1959.1 : Bool;
   "M475" AT %M1959.2 : Bool;
   "M476" AT %M1959.3 : Bool;
   "M477" AT %M1959.4 : Bool;
   "M478" AT %M1959.5 : Bool;
   "M479" AT %M1959.6 : Bool;
   "M480" AT %M1959.7 : Bool;
   "M481" AT %M1960.0 : Bool;
   "M482" AT %M1960.1 : Bool;
   "M483" AT %M1960.2 : Bool;
   "M484" AT %M1960.3 : Bool;
   "M485" AT %M1960.4 : Bool;
   "M486" AT %M1960.5 : Bool;
   "M487" AT %M1960.6 : Bool;
   "M488" AT %M1960.7 : Bool;
   "M489" AT %M1961.0 : Bool;
   "M490" AT %M1961.1 : Bool;
   "M491" AT %M1961.2 : Bool;
   "M492" AT %M1961.3 : Bool;
   "M493" AT %M1961.4 : Bool;
   "M494" AT %M1961.5 : Bool;
   "M495" AT %M1961.6 : Bool;
   "M496" AT %M1961.7 : Bool;
   "M497" AT %M1962.0 : Bool;
   "M498" AT %M1962.1 : Bool;
   "M499" AT %M1962.2 : Bool;
   "M500" AT %M1962.3 : Bool;
   "M501" AT %M1962.4 : Bool;
   "M502" AT %M1962.5 : Bool;
   "M503" AT %M1962.6 : Bool;
   "M504" AT %M1962.7 : Bool;
   "M505" AT %M1963.0 : Bool;
   "M506" AT %M1963.1 : Bool;
   "M507" AT %M1963.2 : Bool;
   "M508" AT %M1963.3 : Bool;
   "M509" AT %M1963.4 : Bool;
   "M510" AT %M1963.5 : Bool;
   "M511" AT %M1963.6 : Bool;
   "M512" AT %M1963.7 : Bool;
   "M513" AT %M1964.0 : Bool;
   "M514" AT %M1964.1 : Bool;
   "M515" AT %M1964.2 : Bool;
   "M516" AT %M1964.3 : Bool;
   "M517" AT %M1964.4 : Bool;
   "M518" AT %M1964.5 : Bool;
   "M519" AT %M1964.6 : Bool;
   "M520" AT %M1964.7 : Bool;
   "Barcode1" AT %MW2000 : Word;
   "Barcode2" AT %MW2002 : Word;
   "Barcode3" AT %MW2004 : Word;
   "Barcode4" AT %MW2006 : Word;
   "Barcode5" AT %MW2008 : Word;
   "Barcode6" AT %MW2010 : Word;
   "Barcode7" AT %MW2012 : Word;
   "Barcode8" AT %MW2014 : Word;
   "Barcode9" AT %MW2016 : Word;
   "Barcode10" AT %MW2018 : Word;
   "Barcode11" AT %MW2020 : Word;
   "Barcode12" AT %MW2022 : Word;
   "Barcode13" AT %MW2024 : Word;
   "Barcode14" AT %MW2026 : Word;
   "Barcode15" AT %MW2028 : Word;
   "Barcode16" AT %MW2030 : Word;
   "Barcode17" AT %MW2032 : Word;
   "Barcode18" AT %MW2034 : Word;
   "Barcode19" AT %MW2036 : Word;
   "Barcode20" AT %MW2038 : Word;
   "Barcode21" AT %MW2040 : Word;
   "Barcode22" AT %MW2042 : Word;
   "Barcode23" AT %MW2044 : Word;
   "Barcode24" AT %MW2046 : Word;
   "Barcode25" AT %MW2048 : Word;
   "Barcode26" AT %MW2050 : Word;
   "Barcode27" AT %MW2052 : Word;
   "Barcode28" AT %MW2054 : Word;
   "Barcode29" AT %MW2056 : Word;
   "Barcode30" AT %MW2058 : Word;
   "Barcode31" AT %MW2060 : Word;
   "Barcode32" AT %MW2062 : Word;
   "Barcode33" AT %MW2064 : Word;
   "Barcode34" AT %MW2066 : Word;
   "Barcode35" AT %MW2068 : Word;
   "Barcode36" AT %MW2070 : Word;
   "Barcode37" AT %MW2072 : Word;
   "Barcode38" AT %MW2074 : Word;
   "Barcode39" AT %MW2076 : Word;
   "Barcode40" AT %MW2078 : Word;
   "Barcode41" AT %MW2080 : Word;
   "Barcode42" AT %MW2082 : Word;
   "Barcode43" AT %MW2084 : Word;
   "Barcode44" AT %MW2086 : Word;
   "Barcode45" AT %MW2088 : Word;
   "Barcode46" AT %MW2090 : Word;
   "Barcode47" AT %MW2092 : Word;
   "Barcode48" AT %MW2094 : Word;
   "Barcode49" AT %MW2096 : Word;
   "Barcode50" AT %MW2098 : Word;
   "Barcode51" AT %MW2100 : Word;
   "Barcode52" AT %MW2102 : Word;
   "Barcode53" AT %MW2104 : Word;
   "Barcode54" AT %MW2106 : Word;
   "Barcode55" AT %MW2108 : Word;
   "Barcode56" AT %MW2110 : Word;
   "Barcode57" AT %MW2112 : Word;
   "Barcode58" AT %MW2114 : Word;
   "Barcode59" AT %MW2116 : Word;
   "Barcode60" AT %MW2118 : Word;
   "Barcode61" AT %MW2120 : Word;
   "Barcode62" AT %MW2122 : Word;
   "Barcode63" AT %MW2124 : Word;
   "Barcode64" AT %MW2126 : Word;
   "Barcode65" AT %MW2128 : Word;
   "Barcode66" AT %MW2130 : Word;
   "Barcode67" AT %MW2132 : Word;
   "Barcode68" AT %MW2134 : Word;
   "Barcode69" AT %MW2136 : Word;
   "Barcode70" AT %MW2138 : Word;
   "Barcode71" AT %MW2140 : Word;
   "Barcode72" AT %MW2142 : Word;
   "Barcode73" AT %MW2144 : Word;
   "Barcode74" AT %MW2146 : Word;
   "Barcode75" AT %MW2148 : Word;
   "Barcode76" AT %MW2150 : Word;
   "Barcode77" AT %MW2152 : Word;
   "Barcode78" AT %MW2154 : Word;
   "Barcode79" AT %MW2156 : Word;
   "Barcode80" AT %MW2158 : Word;
   "Barcode81" AT %MW2160 : Word;
   "Barcode82" AT %MW2162 : Word;
   "Barcode83" AT %MW2164 : Word;
   "Barcode84" AT %MW2166 : Word;
   "Barcode85" AT %MW2168 : Word;
   "Barcode86" AT %MW2170 : Word;
   "Barcode87" AT %MW2172 : Word;
   "Barcode88" AT %MW2174 : Word;
   "Barcode89" AT %MW2176 : Word;
   "Barcode90" AT %MW2178 : Word;
   "Barcode91" AT %MW2180 : Word;
   "Barcode92" AT %MW2182 : Word;
   "Barcode93" AT %MW2184 : Word;
   "Barcode94" AT %MW2186 : Word;
   "Barcode95" AT %MW2188 : Word;
   "Barcode96" AT %MW2190 : Word;
   "Barcode97" AT %MW2192 : Word;
   "Barcode98" AT %MW2194 : Word;
   "Barcode99" AT %MW2196 : Word;
   "Barcode100" AT %MW2198 : Word;
   "Barcode101" AT %MW2200 : Word;
   "Barcode102" AT %MW2202 : Word;
   "Barcode103" AT %MW2204 : Word;
   "Barcode104" AT %MW2206 : Word;
   "Barcode105" AT %MW2208 : Word;
   "Barcode106" AT %MW2210 : Word;
   "Barcode107" AT %MW2212 : Word;
   "Barcode108" AT %MW2214 : Word;
   "Barcode109" AT %MW2216 : Word;
   "Barcode110" AT %MW2218 : Word;
   "Barcode111" AT %MW2220 : Word;
   "Barcode112" AT %MW2222 : Word;
   "Barcode113" AT %MW2224 : Word;
   "Barcode114" AT %MW2226 : Word;
   "Barcode115" AT %MW2228 : Word;
   "Barcode116" AT %MW2230 : Word;
   "Barcode117" AT %MW2232 : Word;
   "Barcode118" AT %MW2234 : Word;
   "Barcode119" AT %MW2236 : Word;
   "Barcode120" AT %MW2238 : Word;
   "Barcode121" AT %MW2240 : Word;
   "Barcode122" AT %MW2242 : Word;
   "Barcode123" AT %MW2244 : Word;
   "Barcode124" AT %MW2246 : Word;
   "Barcode125" AT %MW2248 : Word;
   "Barcode126" AT %MW2250 : Word;
   "Barcode127" AT %MW2252 : Word;
   "Barcode128" AT %MW2254 : Word;
   "Barcode129" AT %MW2256 : Word;
   "Barcode130" AT %MW2258 : Word;
   "Barcode131" AT %MW2260 : Word;
   "Barcode132" AT %MW2262 : Word;
   "Barcode133" AT %MW2264 : Word;
   "Barcode134" AT %MW2266 : Word;
   "Barcode135" AT %MW2268 : Word;
   "Barcode136" AT %MW2270 : Word;
   "Barcode137" AT %MW2272 : Word;
   "Barcode138" AT %MW2274 : Word;
   "Barcode139" AT %MW2276 : Word;
   "Barcode140" AT %MW2278 : Word;
   "Barcode141" AT %MW2280 : Word;
   "Barcode142" AT %MW2282 : Word;
   "Barcode143" AT %MW2284 : Word;
   "Barcode144" AT %MW2286 : Word;
   "Barcode145" AT %MW2288 : Word;
   "Barcode146" AT %MW2290 : Word;
   "Barcode147" AT %MW2292 : Word;
   "Barcode148" AT %MW2294 : Word;
   "Barcode149" AT %MW2296 : Word;
   "Barcode150" AT %MW2298 : Word;
   "Barcode151" AT %MW2300 : Word;
   "Barcode152" AT %MW2302 : Word;
   "Barcode153" AT %MW2304 : Word;
   "Barcode154" AT %MW2306 : Word;
   "Barcode155" AT %MW2308 : Word;
   "Barcode156" AT %MW2310 : Word;
   "Barcode157" AT %MW2312 : Word;
   "Barcode158" AT %MW2314 : Word;
   "Barcode159" AT %MW2316 : Word;
   "Barcode160" AT %MW2318 : Word;
   "Barcode161" AT %MW2320 : Word;
   "Barcode162" AT %MW2322 : Word;
   "Barcode163" AT %MW2324 : Word;
   "Barcode164" AT %MW2326 : Word;
   "Barcode165" AT %MW2328 : Word;
   "Barcode166" AT %MW2330 : Word;
   "Barcode167" AT %MW2332 : Word;
   "Barcode168" AT %MW2334 : Word;
   "Barcode169" AT %MW2336 : Word;
   "Barcode170" AT %MW2338 : Word;
   "Barcode171" AT %MW2340 : Word;
   "Barcode172" AT %MW2342 : Word;
   "Barcode173" AT %MW2344 : Word;
   "Barcode174" AT %MW2346 : Word;
   "Barcode175" AT %MW2348 : Word;
   "Barcode176" AT %MW2350 : Word;
   "Barcode177" AT %MW2352 : Word;
   "Barcode178" AT %MW2354 : Word;
   "Barcode179" AT %MW2356 : Word;
   "Barcode180" AT %MW2358 : Word;
   "Barcode181" AT %MW2360 : Word;
   "Barcode182" AT %MW2362 : Word;
   "Barcode183" AT %MW2364 : Word;
   "Barcode184" AT %MW2366 : Word;
   "Barcode185" AT %MW2368 : Word;
   "Barcode186" AT %MW2370 : Word;
   "Barcode187" AT %MW2372 : Word;
   "Barcode188" AT %MW2374 : Word;
   "Barcode189" AT %MW2376 : Word;
   "Barcode190" AT %MW2378 : Word;
   "Barcode191" AT %MW2380 : Word;
   "Barcode192" AT %MW2382 : Word;
   "Barcode193" AT %MW2384 : Word;
   "Barcode194" AT %MW2386 : Word;
   "Barcode195" AT %MW2388 : Word;
   "Barcode196" AT %MW2390 : Word;
   "Barcode197" AT %MW2392 : Word;
   "Barcode198" AT %MW2394 : Word;
   "Barcode199" AT %MW2396 : Word;
   "Barcode200" AT %MW2398 : Word;
   "Barcode201" AT %MW2400 : Word;
   "Barcode202" AT %MW2402 : Word;
   "Barcode203" AT %MW2404 : Word;
   "Barcode204" AT %MW2406 : Word;
   "Barcode205" AT %MW2408 : Word;
   "Barcode206" AT %MW2410 : Word;
   "Barcode207" AT %MW2412 : Word;
   "Barcode208" AT %MW2414 : Word;
   "Barcode209" AT %MW2416 : Word;
   "Barcode210" AT %MW2418 : Word;
   "Barcode211" AT %MW2420 : Word;
   "Barcode212" AT %MW2422 : Word;
   "Barcode213" AT %MW2424 : Word;
   "Barcode214" AT %MW2426 : Word;
   "Barcode215" AT %MW2428 : Word;
   "Barcode216" AT %MW2430 : Word;
   "Barcode217" AT %MW2432 : Word;
   "Barcode218" AT %MW2434 : Word;
   "Barcode219" AT %MW2436 : Word;
   "Barcode220" AT %MW2438 : Word;
   "Barcode221" AT %MW2440 : Word;
   "Barcode222" AT %MW2442 : Word;
   "Barcode223" AT %MW2444 : Word;
   "Barcode224" AT %MW2446 : Word;
   "Barcode225" AT %MW2448 : Word;
   "Barcode226" AT %MW2450 : Word;
   "Barcode227" AT %MW2452 : Word;
   "Barcode228" AT %MW2454 : Word;
   "Barcode229" AT %MW2456 : Word;
   "Barcode230" AT %MW2458 : Word;
   "Barcode231" AT %MW2460 : Word;
   "Barcode232" AT %MW2462 : Word;
   "Barcode233" AT %MW2464 : Word;
   "Barcode234" AT %MW2466 : Word;
   "Barcode235" AT %MW2468 : Word;
   "Barcode236" AT %MW2470 : Word;
   "Barcode237" AT %MW2472 : Word;
   "Barcode238" AT %MW2474 : Word;
   "Barcode239" AT %MW2476 : Word;
   "Barcode240" AT %MW2478 : Word;
   "Barcode241" AT %MW2480 : Word;
   "Barcode242" AT %MW2482 : Word;
   "Barcode243" AT %MW2484 : Word;
   "Barcode244" AT %MW2486 : Word;
   "Barcode245" AT %MW2488 : Word;
   "Barcode246" AT %MW2490 : Word;
   "Barcode247" AT %MW2492 : Word;
   "Barcode248" AT %MW2494 : Word;
   "Barcode249" AT %MW2496 : Word;
   "Barcode250" AT %MW2498 : Word;
   "Barcode251" AT %MW2500 : Word;
   "Barcode252" AT %MW2502 : Word;
   "Barcode253" AT %MW2504 : Word;
   "Barcode254" AT %MW2506 : Word;
   "Barcode255" AT %MW2508 : Word;
   "Barcode256" AT %MW2510 : Word;
   "Barcode257" AT %MW2512 : Word;
   "Barcode258" AT %MW2514 : Word;
   "Barcode259" AT %MW2516 : Word;
   "Barcode260" AT %MW2518 : Word;
   "Barcode261" AT %MW2520 : Word;
   "Barcode262" AT %MW2522 : Word;
   "Barcode263" AT %MW2524 : Word;
   "Barcode264" AT %MW2526 : Word;
   "Barcode265" AT %MW2528 : Word;
   "Barcode266" AT %MW2530 : Word;
   "Barcode267" AT %MW2532 : Word;
   "Barcode268" AT %MW2534 : Word;
   "Barcode269" AT %MW2536 : Word;
   "Barcode270" AT %MW2538 : Word;
   "Barcode271" AT %MW2540 : Word;
   "Barcode272" AT %MW2542 : Word;
   "Barcode273" AT %MW2544 : Word;
   "Barcode274" AT %MW2546 : Word;
   "Barcode275" AT %MW2548 : Word;
   "Barcode276" AT %MW2550 : Word;
   "Barcode277" AT %MW2552 : Word;
   "Barcode278" AT %MW2554 : Word;
   "Barcode279" AT %MW2556 : Word;
   "Barcode280" AT %MW2558 : Word;
   "Barcode281" AT %MW2560 : Word;
   "Barcode282" AT %MW2562 : Word;
   "Barcode283" AT %MW2564 : Word;
   "Barcode284" AT %MW2566 : Word;
   "Barcode285" AT %MW2568 : Word;
   "Barcode286" AT %MW2570 : Word;
   "Barcode287" AT %MW2572 : Word;
   "Barcode288" AT %MW2574 : Word;
   "Barcode289" AT %MW2576 : Word;
   "Barcode290" AT %MW2578 : Word;
   "Barcode291" AT %MW2580 : Word;
   "Barcode292" AT %MW2582 : Word;
   "Barcode293" AT %MW2584 : Word;
   "Barcode294" AT %MW2586 : Word;
   "Barcode295" AT %MW2588 : Word;
   "Barcode296" AT %MW2590 : Word;
   "Barcode297" AT %MW2592 : Word;
   "Barcode298" AT %MW2594 : Word;
   "Barcode299" AT %MW2596 : Word;
   "Barcode300" AT %MW2598 : Word;
   "Barcode301" AT %MW2600 : Word;
   "Barcode302" AT %MW2602 : Word;
   "Barcode303" AT %MW2604 : Word;
   "Barcode304" AT %MW2606 : Word;
   "Barcode305" AT %MW2608 : Word;
   "Barcode306" AT %MW2610 : Word;
   "Barcode307" AT %MW2612 : Word;
   "Barcode308" AT %MW2614 : Word;
   "Barcode309" AT %MW2616 : Word;
   "Barcode310" AT %MW2618 : Word;
   "Barcode311" AT %MW2620 : Word;
   "Barcode312" AT %MW2622 : Word;
   "Barcode313" AT %MW2624 : Word;
   "Barcode314" AT %MW2626 : Word;
   "Barcode315" AT %MW2628 : Word;
   "Barcode316" AT %MW2630 : Word;
   "Barcode317" AT %MW2632 : Word;
   "Barcode318" AT %MW2634 : Word;
   "Barcode319" AT %MW2636 : Word;
   "Barcode320" AT %MW2638 : Word;
   "Barcode321" AT %MW2640 : Word;
   "Barcode322" AT %MW2642 : Word;
   "Barcode323" AT %MW2644 : Word;
   "Barcode324" AT %MW2646 : Word;
   "Barcode325" AT %MW2648 : Word;
   "Barcode326" AT %MW2650 : Word;
   "Barcode327" AT %MW2652 : Word;
   "Barcode328" AT %MW2654 : Word;
   "Barcode329" AT %MW2656 : Word;
   "Barcode330" AT %MW2658 : Word;
   "Barcode331" AT %MW2660 : Word;
   "Barcode332" AT %MW2662 : Word;
   "Barcode333" AT %MW2664 : Word;
   "Barcode334" AT %MW2666 : Word;
   "Barcode335" AT %MW2668 : Word;
   "Barcode336" AT %MW2670 : Word;
   "Barcode337" AT %MW2672 : Word;
   "Barcode338" AT %MW2674 : Word;
   "Barcode339" AT %MW2676 : Word;
   "Barcode340" AT %MW2678 : Word;
   "Barcode341" AT %MW2680 : Word;
   "Barcode342" AT %MW2682 : Word;
   "Barcode343" AT %MW2684 : Word;
   "Barcode344" AT %MW2686 : Word;
   "Barcode345" AT %MW2688 : Word;
   "Barcode346" AT %MW2690 : Word;
   "Barcode347" AT %MW2692 : Word;
   "Barcode348" AT %MW2694 : Word;
   "Barcode349" AT %MW2696 : Word;
   "Barcode350" AT %MW2698 : Word;
   "Barcode351" AT %MW2700 : Word;
   "Barcode352" AT %MW2702 : Word;
   "Barcode353" AT %MW2704 : Word;
   "Barcode354" AT %MW2706 : Word;
   "Barcode355" AT %MW2708 : Word;
   "Barcode356" AT %MW2710 : Word;
   "Barcode357" AT %MW2712 : Word;
   "Barcode358" AT %MW2714 : Word;
   "Barcode359" AT %MW2716 : Word;
   "Barcode360" AT %MW2718 : Word;
   "Barcode361" AT %MW2720 : Word;
   "Barcode362" AT %MW2722 : Word;
   "Barcode363" AT %MW2724 : Word;
   "Barcode364" AT %MW2726 : Word;
   "Barcode365" AT %MW2728 : Word;
   "Barcode366" AT %MW2730 : Word;
   "Barcode367" AT %MW2732 : Word;
   "Barcode368" AT %MW2734 : Word;
   "Barcode369" AT %MW2736 : Word;
   "Barcode370" AT %MW2738 : Word;
   "Barcode371" AT %MW2740 : Word;
   "Barcode372" AT %MW2742 : Word;
   "Barcode373" AT %MW2744 : Word;
   "Barcode374" AT %MW2746 : Word;
   "Barcode375" AT %MW2748 : Word;
   "Barcode376" AT %MW2750 : Word;
   "Barcode377" AT %MW2752 : Word;
   "Barcode378" AT %MW2754 : Word;
   "Barcode379" AT %MW2756 : Word;
   "Barcode380" AT %MW2758 : Word;
   "Barcode381" AT %MW2760 : Word;
   "Barcode382" AT %MW2762 : Word;
   "Barcode383" AT %MW2764 : Word;
   "Barcode384" AT %MW2766 : Word;
   "Barcode385" AT %MW2768 : Word;
   "Barcode386" AT %MW2770 : Word;
   "Barcode387" AT %MW2772 : Word;
   "Barcode388" AT %MW2774 : Word;
   "Barcode389" AT %MW2776 : Word;
   "Barcode390" AT %MW2778 : Word;
   "Barcode391" AT %MW2780 : Word;
   "Barcode392" AT %MW2782 : Word;
   "Barcode393" AT %MW2784 : Word;
   "Barcode394" AT %MW2786 : Word;
   "Barcode395" AT %MW2788 : Word;
   "Barcode396" AT %MW2790 : Word;
   "Barcode397" AT %MW2792 : Word;
   "Barcode398" AT %MW2794 : Word;
   "Barcode399" AT %MW2796 : Word;
   "Barcode400" AT %MW2798 : Word;
   "Barcode401" AT %MW2800 : Word;
   "Barcode402" AT %MW2802 : Word;
   "Barcode403" AT %MW2804 : Word;
   "Barcode404" AT %MW2806 : Word;
   "Barcode405" AT %MW2808 : Word;
   "Barcode406" AT %MW2810 : Word;
   "Barcode407" AT %MW2812 : Word;
   "Barcode408" AT %MW2814 : Word;
   "Barcode409" AT %MW2816 : Word;
   "Barcode410" AT %MW2818 : Word;
   "Barcode411" AT %MW2820 : Word;
   "Barcode412" AT %MW2822 : Word;
   "Barcode413" AT %MW2824 : Word;
   "Barcode414" AT %MW2826 : Word;
   "Barcode415" AT %MW2828 : Word;
   "Barcode416" AT %MW2830 : Word;
   "Barcode417" AT %MW2832 : Word;
   "Barcode418" AT %MW2834 : Word;
   "Barcode419" AT %MW2836 : Word;
   "Barcode420" AT %MW2838 : Word;
   "Barcode421" AT %MW2840 : Word;
   "Barcode422" AT %MW2842 : Word;
   "Barcode423" AT %MW2844 : Word;
   "Barcode424" AT %MW2846 : Word;
   "Barcode425" AT %MW2848 : Word;
   "Barcode426" AT %MW2850 : Word;
   "Barcode427" AT %MW2852 : Word;
   "Barcode428" AT %MW2854 : Word;
   "Barcode429" AT %MW2856 : Word;
   "Barcode430" AT %MW2858 : Word;
   "Barcode431" AT %MW2860 : Word;
   "Barcode432" AT %MW2862 : Word;
   "Barcode433" AT %MW2864 : Word;
   "Barcode434" AT %MW2866 : Word;
   "Barcode435" AT %MW2868 : Word;
   "Barcode436" AT %MW2870 : Word;
   "Barcode437" AT %MW2872 : Word;
   "Barcode438" AT %MW2874 : Word;
   "Barcode439" AT %MW2876 : Word;
   "Barcode440" AT %MW2878 : Word;
   "Barcode441" AT %MW2880 : Word;
   "Barcode442" AT %MW2882 : Word;
   "Barcode443" AT %MW2884 : Word;
   "Barcode444" AT %MW2886 : Word;
   "Barcode445" AT %MW2888 : Word;
   "Barcode446" AT %MW2890 : Word;
   "Barcode447" AT %MW2892 : Word;
   "Barcode448" AT %MW2894 : Word;
   "Barcode449" AT %MW2896 : Word;
   "Barcode450" AT %MW2898 : Word;
   "Barcode451" AT %MW2900 : Word;
   "Barcode452" AT %MW2902 : Word;
   "Barcode453" AT %MW2904 : Word;
   "Barcode454" AT %MW2906 : Word;
   "Barcode455" AT %MW2908 : Word;
   "Barcode456" AT %MW2910 : Word;
   "Barcode457" AT %MW2912 : Word;
   "Barcode458" AT %MW2914 : Word;
   "Barcode459" AT %MW2916 : Word;
   "Barcode460" AT %MW2918 : Word;
   "Barcode461" AT %MW2920 : Word;
   "Barcode462" AT %MW2922 : Word;
   "Barcode463" AT %MW2924 : Word;
   "Barcode464" AT %MW2926 : Word;
   "Barcode465" AT %MW2928 : Word;
   "Barcode466" AT %MW2930 : Word;
   "Barcode467" AT %MW2932 : Word;
   "Barcode468" AT %MW2934 : Word;
   "Barcode469" AT %MW2936 : Word;
   "Barcode470" AT %MW2938 : Word;
   "Barcode471" AT %MW2940 : Word;
   "Barcode472" AT %MW2942 : Word;
   "Barcode473" AT %MW2944 : Word;
   "Barcode474" AT %MW2946 : Word;
   "Barcode475" AT %MW2948 : Word;
   "Barcode476" AT %MW2950 : Word;
   "Barcode477" AT %MW2952 : Word;
   "Barcode478" AT %MW2954 : Word;
   "Barcode479" AT %MW2956 : Word;
   "Barcode480" AT %MW2958 : Word;
   "Barcode481" AT %MW2960 : Word;
   "Barcode482" AT %MW2962 : Word;
   "Barcode483" AT %MW2964 : Word;
   "Barcode484" AT %MW2966 : Word;
   "Barcode485" AT %MW2968 : Word;
   "Barcode486" AT %MW2970 : Word;
   "Barcode487" AT %MW2972 : Word;
   "Barcode488" AT %MW2974 : Word;
   "Barcode489" AT %MW2976 : Word;
   "Barcode490" AT %MW2978 : Word;
   "Barcode491" AT %MW2980 : Word;
   "Barcode492" AT %MW2982 : Word;
   "Barcode493" AT %MW2984 : Word;
   "Barcode494" AT %MW2986 : Word;
   "Barcode495" AT %MW2988 : Word;
   "Barcode496" AT %MW2990 : Word;
   "Barcode497" AT %MW2992 : Word;
   "Barcode498" AT %MW2994 : Word;
   "Barcode499" AT %MW2996 : Word;
   "Barcode500" AT %MW2998 : Word;
   "Barcode501" AT %MW3000 : Word;
   "Barcode502" AT %MW3002 : Word;
   "Barcode503" AT %MW3004 : Word;
   "Barcode504" AT %MW3006 : Word;
   "Barcode505" AT %MW3008 : Word;
   "Barcode506" AT %MW3010 : Word;
   "Barcode507" AT %MW3012 : Word;
   "Barcode508" AT %MW3014 : Word;
   "Barcode509" AT %MW3016 : Word;
   "Barcode510" AT %MW3018 : Word;
   "Barcode511" AT %MW3020 : Word;
   "Barcode512" AT %MW3022 : Word;
   "Barcode513" AT %MW3024 : Word;
   "Barcode514" AT %MW3026 : Word;
   "Barcode515" AT %MW3028 : Word;
   "Barcode516" AT %MW3030 : Word;
   "Barcode517" AT %MW3032 : Word;
   "Barcode518" AT %MW3034 : Word;
   "Barcode519" AT %MW3036 : Word;
   "Barcode520" AT %MW3038 : Word;
   "Button_OK_Screen" AT %M3040.0 : Bool;
   "แสดงชื่อยา" AT %MW3042 : Word;
   "Output Resrt_ชื่อยา" AT %M3500.0 : Bool;
   "ป้อนรหัส Barcode" AT %I100.6 : Bool;
   "Gripper เคลื่อนไปช่องยา" AT %I101.0 : Bool;
   "Gripper วางยา" AT %I101.1 : Bool;
   "เคลื่อนที่ไปยังจุดเริ่มต้น" AT %I101.2 : Bool;
   "รอรับคำสั่งยา" AT %I101.3 : Bool;
   "Gripperเคลื่อนที่มาเอายา" AT %I100.7 : Bool;
   "รับคำสั่งเบิกยา" AT %I101.4 : Bool;
   "เคลื่อนที่ไปยังตำยา" AT %I101.5 : Bool;
   "เคลื่อนที่ไปยังตำแหน่งเริ่มต้น เบิกจ่าย" AT %I101.7 : Bool;
   "รอคำสั่งเบิกยา" AT %I102.0 : Bool;
   "Gripper หยิบยา" AT %I102.1 : Bool;
   "Output Status1" AT %MW3054 : Word;
   "Output Status2" AT %MW3056 : Word;
   "ปุ่มยืนยันหน้า Screen" AT %M1965.0 : Bool;
   "ปุ่มClear" AT %M1965.2 : Bool;
END_VAR

DATA_BLOCK "Step motor ขึ่น-ลง ตามแกน y No.1_Forword_DB"   // DB13
{ S7_Optimized_Access := 'TRUE' }
VERSION : 0.1
// stored: InstanceOfName Step motor ขึ่น-ลง ตามแกน y No.1,No.2_Forword
"Step motor ขึ่น-ลง ตามแกน y No.1,No.2_Forword"
BEGIN
END_DATA_BLOCK

DATA_BLOCK "Step motor ขึ่น-ลง ตามแกน y No.1,No.2_Forword_DB"   // DB22
{ S7_Optimized_Access := 'TRUE' }
VERSION : 0.1
// stored: InstanceOfName Step motor ขึ่น-ลง ตามแกน y No.1,No.2_Forword
"Step motor ขึ่น-ลง ตามแกน y No.1,No.2_Forword"
BEGIN
END_DATA_BLOCK

DATA_BLOCK "Step motor ซ้าน-ขวา ตามแกน X  No.1_Forword_DB"   // DB26
{ S7_Optimized_Access := 'TRUE' }
VERSION : 0.1
// stored: InstanceOfName Step motor ซ้าน-ขวา ตามแกน X No.1_Forword
"Step motor ซ้าน-ขวา ตามแกน X  No.1_Forword"
BEGIN
END_DATA_BLOCK

DATA_BLOCK "Step motor ขึ่น-ลง ตามแกน y No.1,No.2_Blackword_DB"   // DB29
{ S7_Optimized_Access := 'TRUE' }
VERSION : 0.1
// stored: InstanceOfName Step motor ขึ่น-ลง ตามแกน y No.1_Blackword
"Step motor ขึ่น-ลง ตามแกน y No.1_Blackword"
BEGIN
END_DATA_BLOCK

DATA_BLOCK "Gripper_DB"   // DB64
{ S7_Optimized_Access := 'TRUE' }
VERSION : 0.1
// stored: InstanceOfName Gripper
"Gripper"
BEGIN
END_DATA_BLOCK

DATA_BLOCK "Step motor ซ้าย-ขวา ตามแกน X No.1_Blackword_DB"   // DB66
{ S7_Optimized_Access := 'TRUE' }
VERSION : 0.1
// stored: InstanceOfName Step motor ซ้าย-ขวา ตามแกน X No.1_Blackword
"Step motor ซ้าย-ขวา ตามแกน X No.1_Blackword"
BEGIN
END_DATA_BLOCK

DATA_BLOCK "Step motor ขึ่น-ลง ตามแกน y No.1,No.2_Forword(เบิกจ่าย)_DB"   // DB152
{ S7_Optimized_Access := 'TRUE' }
VERSION : 0.1
// stored: InstanceOfName Step motor ขึ่น-ลง ตามแกน y No.1,No.2_Forword(เบิกจ่าย)
"Step motor ขึ่น-ลง ตามแกน y No.1,No.2_Forword(เบิกจ่าย)"
BEGIN
END_DATA_BLOCK

DATA_BLOCK "Step motor ขึ่น-ลง ตามแกน y No.1,No.2_Blackword(เบิกจ่าย)_DB"   // DB173
{ S7_Optimized_Access := 'TRUE' }
VERSION : 0.1
// stored: InstanceOfName Step motor ขึ่น-ลง ตามแกน y No.1,No.2_Blackword(เบิกจ่าย)
"Step motor ขึ่น-ลง ตามแกน y No.1,No.2_Blackword(เบิกจ่าย)"
BEGIN
END_DATA_BLOCK

DATA_BLOCK "Gripper_เบิกจ่าย_DB"   // DB174
{ S7_Optimized_Access := 'TRUE' }
VERSION : 0.1
// stored: InstanceOfName Gripper_เบิกจ่าย
"Gripper_เบิกจ่าย"
BEGIN
END_DATA_BLOCK

DATA_BLOCK "Step motor ขึ่น-ลง ตามแกน y No.3_Forword(เบิกจ่าย)_DB"   // DB229
{ S7_Optimized_Access := 'TRUE' }
VERSION : 0.1
// stored: InstanceOfName Step motor ขึ่น-ลง ตามแกน y No.3_Forword(เบิกจ่าย)
"Step motor ขึ่น-ลง ตามแกน y No.3_Forword(เบิกจ่าย)"
BEGIN
END_DATA_BLOCK

DATA_BLOCK "Step motor ขึ่น-ลง ตามแกน y No.3_Blackword(เบิกจ่าย)_DB"   // DB230
{ S7_Optimized_Access := 'TRUE' }
VERSION : 0.1
// stored: InstanceOfName Step motor ขึ่น-ลง ตามแกน y No.3_Blackword(เบิกจ่าย)
"Step motor ขึ่น-ลง ตามแกน y No.3_Blackword(เบิกจ่าย)"
BEGIN
END_DATA_BLOCK

DATA_BLOCK "บันทึกผลการเคลื่อนที่ ไว้ที่ Excell_DB"   // DB235
{ S7_Optimized_Access := 'TRUE' }
VERSION : 0.1
// stored: InstanceOfName บันทึกผลการเคลื่อนที่ ไว้ที่ Excell
"บันทึกผลการเคลื่อนที่ ไว้ที่ Excell"
BEGIN
END_DATA_BLOCK

DATA_BLOCK "Screen Data Pro จัดเก็บ_DB"   // DB758
{ S7_Optimized_Access := 'TRUE' }
VERSION : 0.1
// stored: InstanceOfName Screen Data Pro จัดเก็บ
"Screen Data Pro จัดเก็บ"
BEGIN
END_DATA_BLOCK

// folder: System blocks/Program resources

DATA_BLOCK "IEC_Timer_0_DB"   // DB1
{ S7_Optimized_Access := 'TRUE' }
AUTHOR : Simatic
FAMILY : IEC
NAME : IEC_TMR
VERSION : 1.0
// stored: InstanceOfName IEC_TIMER
"IEC_TIMER"
BEGIN
END_DATA_BLOCK

DATA_BLOCK "Timer_1"   // DB3
{ S7_Optimized_Access := 'TRUE' }
AUTHOR : Simatic
FAMILY : IEC
NAME : IEC_TMR
VERSION : 1.0
// stored: InstanceOfName IEC_TIMER
"IEC_TIMER"
BEGIN
END_DATA_BLOCK

DATA_BLOCK "Timer_2"   // DB4
{ S7_Optimized_Access := 'TRUE' }
AUTHOR : Simatic
FAMILY : IEC
NAME : IEC_TMR
VERSION : 1.0
// stored: InstanceOfName IEC_TIMER
"IEC_TIMER"
BEGIN
END_DATA_BLOCK

DATA_BLOCK "Timer_3"   // DB5
{ S7_Optimized_Access := 'TRUE' }
AUTHOR : Simatic
FAMILY : IEC
NAME : IEC_TMR
VERSION : 1.0
// stored: InstanceOfName IEC_TIMER
"IEC_TIMER"
BEGIN
END_DATA_BLOCK

DATA_BLOCK "Timer_4"   // DB6
{ S7_Optimized_Access := 'TRUE' }
AUTHOR : Simatic
FAMILY : IEC
NAME : IEC_TMR
VERSION : 1.0
// stored: InstanceOfName IEC_TIMER
"IEC_TIMER"
BEGIN
END_DATA_BLOCK

DATA_BLOCK "Timer_5"   // DB7
{ S7_Optimized_Access := 'TRUE' }
AUTHOR : Simatic
FAMILY : IEC
NAME : IEC_TMR
VERSION : 1.0
// stored: InstanceOfName IEC_TIMER
"IEC_TIMER"
BEGIN
END_DATA_BLOCK

DATA_BLOCK "Timer_6"   // DB8
{ S7_Optimized_Access := 'TRUE' }
AUTHOR : Simatic
FAMILY : IEC
NAME : IEC_TMR
VERSION : 1.0
// stored: InstanceOfName IEC_TIMER
"IEC_TIMER"
BEGIN
END_DATA_BLOCK

DATA_BLOCK "Timer_7"   // DB9
{ S7_Optimized_Access := 'TRUE' }
AUTHOR : Simatic
FAMILY : IEC
NAME : IEC_TMR
VERSION : 1.0
// stored: InstanceOfName IEC_TIMER
"IEC_TIMER"
BEGIN
END_DATA_BLOCK

DATA_BLOCK "Timer_8"   // DB10
{ S7_Optimized_Access := 'TRUE' }
AUTHOR : Simatic
FAMILY : IEC
NAME : IEC_TMR
VERSION : 1.0
// stored: InstanceOfName IEC_TIMER
"IEC_TIMER"
BEGIN
END_DATA_BLOCK

DATA_BLOCK "Timer_9"   // DB11
{ S7_Optimized_Access := 'TRUE' }
AUTHOR : Simatic
FAMILY : IEC
NAME : IEC_TMR
VERSION : 1.0
// stored: InstanceOfName IEC_TIMER
"IEC_TIMER"
BEGIN
END_DATA_BLOCK

DATA_BLOCK "Timer_10"   // DB12
{ S7_Optimized_Access := 'TRUE' }
AUTHOR : Simatic
FAMILY : IEC
NAME : IEC_TMR
VERSION : 1.0
// stored: InstanceOfName IEC_TIMER
"IEC_TIMER"
BEGIN
END_DATA_BLOCK

DATA_BLOCK "Timer_11"   // DB14
{ S7_Optimized_Access := 'TRUE' }
AUTHOR : Simatic
FAMILY : IEC
NAME : IEC_TMR
VERSION : 1.0
// stored: InstanceOfName IEC_TIMER
"IEC_TIMER"
BEGIN
END_DATA_BLOCK

DATA_BLOCK "Timer_12"   // DB15
{ S7_Optimized_Access := 'TRUE' }
AUTHOR : Simatic
FAMILY : IEC
NAME : IEC_TMR
VERSION : 1.0
// stored: InstanceOfName IEC_TIMER
"IEC_TIMER"
BEGIN
END_DATA_BLOCK

DATA_BLOCK "Timer_13"   // DB16
{ S7_Optimized_Access := 'TRUE' }
AUTHOR : Simatic
FAMILY : IEC
NAME : IEC_TMR
VERSION : 1.0
// stored: InstanceOfName IEC_TIMER
"IEC_TIMER"
BEGIN
END_DATA_BLOCK

DATA_BLOCK "Timer_14"   // DB17
{ S7_Optimized_Access := 'TRUE' }
AUTHOR : Simatic
FAMILY : IEC
NAME : IEC_TMR
VERSION : 1.0
// stored: InstanceOfName IEC_TIMER
"IEC_TIMER"
BEGIN
END_DATA_BLOCK

DATA_BLOCK "Timer_16"   // DB18
{ S7_Optimized_Access := 'TRUE' }
AUTHOR : Simatic
FAMILY : IEC
NAME : IEC_TMR
VERSION : 1.0
// stored: InstanceOfName IEC_TIMER
"IEC_TIMER"
BEGIN
END_DATA_BLOCK

DATA_BLOCK "Timer_15"   // DB19
{ S7_Optimized_Access := 'TRUE' }
AUTHOR : Simatic
FAMILY : IEC
NAME : IEC_TMR
VERSION : 1.0
// stored: InstanceOfName IEC_TIMER
"IEC_TIMER"
BEGIN
END_DATA_BLOCK

DATA_BLOCK "Timer_17"   // DB20
{ S7_Optimized_Access := 'TRUE' }
AUTHOR : Simatic
FAMILY : IEC
NAME : IEC_TMR
VERSION : 1.0
// stored: InstanceOfName IEC_TIMER
"IEC_TIMER"
BEGIN
END_DATA_BLOCK

DATA_BLOCK "Timer_18"   // DB21
{ S7_Optimized_Access := 'TRUE' }
AUTHOR : Simatic
FAMILY : IEC
NAME : IEC_TMR
VERSION : 1.0
// stored: InstanceOfName IEC_TIMER
"IEC_TIMER"
BEGIN
END_DATA_BLOCK

DATA_BLOCK "Timer_19"   // DB23
{ S7_Optimized_Access := 'TRUE' }
AUTHOR : Simatic
FAMILY : IEC
NAME : IEC_TMR
VERSION : 1.0
// stored: InstanceOfName IEC_TIMER
"IEC_TIMER"
BEGIN
END_DATA_BLOCK

DATA_BLOCK "Timer_20"   // DB24
{ S7_Optimized_Access := 'TRUE' }
AUTHOR : Simatic
FAMILY : IEC
NAME : IEC_TMR
VERSION : 1.0
// stored: InstanceOfName IEC_TIMER
"IEC_TIMER"
BEGIN
END_DATA_BLOCK

DATA_BLOCK "IEC_Timer_0_DB_1"   // DB25
{ S7_Optimized_Access := 'TRUE' }
AUTHOR : Simatic
FAMILY : IEC
NAME : IEC_TMR
VERSION : 1.0
// stored: InstanceOfName IEC_TIMER
"IEC_TIMER"
BEGIN
END_DATA_BLOCK

DATA_BLOCK "IEC_Timer_0_DB_2"   // DB28
{ S7_Optimized_Access := 'TRUE' }
AUTHOR : Simatic
FAMILY : IEC
NAME : IEC_TMR
VERSION : 1.0
// stored: InstanceOfName IEC_TIMER
"IEC_TIMER"
BEGIN
END_DATA_BLOCK

DATA_BLOCK "IEC_Timer_0_DB_4"   // DB30
{ S7_Optimized_Access := 'TRUE' }
AUTHOR : Simatic
FAMILY : IEC
NAME : IEC_TMR
VERSION : 1.0
// stored: InstanceOfName IEC_TIMER
"IEC_TIMER"
BEGIN
END_DATA_BLOCK

DATA_BLOCK "IEC_Timer_0_DB_5"   // DB31
{ S7_Optimized_Access := 'TRUE' }
AUTHOR : Simatic
FAMILY : IEC
NAME : IEC_TMR
VERSION : 1.0
// stored: InstanceOfName IEC_TIMER
"IEC_TIMER"
BEGIN
END_DATA_BLOCK

DATA_BLOCK "IEC_Timer_0_DB_6"   // DB32
{ S7_Optimized_Access := 'TRUE' }
AUTHOR : Simatic
FAMILY : IEC
NAME : IEC_TMR
VERSION : 1.0
// stored: InstanceOfName IEC_TIMER
"IEC_TIMER"
BEGIN
END_DATA_BLOCK

DATA_BLOCK "IEC_Timer_0_DB_7"   // DB33
{ S7_Optimized_Access := 'TRUE' }
AUTHOR : Simatic
FAMILY : IEC
NAME : IEC_TMR
VERSION : 1.0
// stored: InstanceOfName IEC_TIMER
"IEC_TIMER"
BEGIN
END_DATA_BLOCK

DATA_BLOCK "IEC_Timer_0_DB_8"   // DB34
{ S7_Optimized_Access := 'TRUE' }
AUTHOR : Simatic
FAMILY : IEC
NAME : IEC_TMR
VERSION : 1.0
// stored: InstanceOfName IEC_TIMER
"IEC_TIMER"
BEGIN
END_DATA_BLOCK

DATA_BLOCK "IEC_Timer_0_DB_9"   // DB35
{ S7_Optimized_Access := 'TRUE' }
AUTHOR : Simatic
FAMILY : IEC
NAME : IEC_TMR
VERSION : 1.0
// stored: InstanceOfName IEC_TIMER
"IEC_TIMER"
BEGIN
END_DATA_BLOCK

DATA_BLOCK "IEC_Timer_0_DB_10"   // DB36
{ S7_Optimized_Access := 'TRUE' }
AUTHOR : Simatic
FAMILY : IEC
NAME : IEC_TMR
VERSION : 1.0
// stored: InstanceOfName IEC_TIMER
"IEC_TIMER"
BEGIN
END_DATA_BLOCK

DATA_BLOCK "IEC_Timer_0_DB_11"   // DB37
{ S7_Optimized_Access := 'TRUE' }
AUTHOR : Simatic
FAMILY : IEC
NAME : IEC_TMR
VERSION : 1.0
// stored: InstanceOfName IEC_TIMER
"IEC_TIMER"
BEGIN
END_DATA_BLOCK

DATA_BLOCK "IEC_Timer_0_DB_12"   // DB38
{ S7_Optimized_Access := 'TRUE' }
AUTHOR : Simatic
FAMILY : IEC
NAME : IEC_TMR
VERSION : 1.0
// stored: InstanceOfName IEC_TIMER
"IEC_TIMER"
BEGIN
END_DATA_BLOCK

DATA_BLOCK "IEC_Timer_0_DB_13"   // DB39
{ S7_Optimized_Access := 'TRUE' }
AUTHOR : Simatic
FAMILY : IEC
NAME : IEC_TMR
VERSION : 1.0
// stored: InstanceOfName IEC_TIMER
"IEC_TIMER"
BEGIN
END_DATA_BLOCK

